(* IEC 61131-3 sources: volt/packages/volt-lsp-iec/test-corpus/awa-palletizer/Device/Plc Logic/Application/Library Manager/L_TW2P_TechModulesWindingTraversing, 72 files *)

(* ---- L_TW2P_ADAPTSPDCTRLGAINMODE.dut ---- *)
TYPE L_TW2P_ADAPTSPDCTRLGAINMODE :
(
	DIAMTOSQUARE := 0,
	DIAM := 1,
	INERTIA := 2
);
END_TYPE

(* ---- L_TW2P_DANCERCTRLSTOPMODE.dut ---- *)
TYPE L_TW2P_DANCERCTRLSTOPMODE :
(
	HALT := 0,
	MOVEABS := 1,
	MOVEREL := 2,
	MOVEABSSHORTESTWAY := 3,
	STOPVELOCITYMASTER := 4
);
END_TYPE

(* ---- L_TW2P_DANCERLIMITMODE.dut ---- *)
TYPE L_TW2P_DANCERLIMITMODE :
(
	AUTOMATIC := 0,
	SCPARDANCERLIMITS := 1,
	TEACHEDDANCERLIMITS := 2
);
END_TYPE

(* ---- L_TW2P_PERSISTENTVARWINDER.dut ---- *)
TYPE L_TW2P_PERSISTENTVARWINDER :
STRUCT
	LRDIAM : LREAL;
	LRMATERIALCOUNTER : LREAL;
	LIREVCOUNTER : LINT;
	LRREVCOUNTERRESIDUAL : LREAL;
	XUPPERPOSTEACHED : BOOL;
	XLOWERPOSTEACHED : BOOL;
	LRDANCERUPPERLIMIT : LREAL;
	LRDANCERLOWERLIMIT : LREAL;
END_STRUCT
END_TYPE

(* ---- L_TW2P_RESETICTRLMODE.dut ---- *)
TYPE L_TW2P_RESETICTRLMODE :
(
	INSTANT := 0,
	RAMP := 1
);
END_TYPE

(* ---- L_TW2P_SCAP_TM_WINDER.dut ---- *)
TYPE L_TW2P_SCAP_TM_WINDER :
STRUCT
	AP_XSETVELOFFSET : BOOL;
	AP_LRVELOFFSET : LREAL;
	AP_XSETTRQOFFSET : BOOL;
	AP_LRSETTRQOFFSET : LREAL;
	AP_XSETVELOFFSETDIAMCACL : BOOL;
	AP_LRVELOFFSETDIAMCACL : LREAL;
	AP_XSETSPEEDPOINTDIAMCALC : BOOL;
	AP_LRSETSPEEDPOINTDIAMCALC : LREAL;
	AP_XSETSPEEDPOINT : BOOL;
	AP_LRSETSPEEDPOINT : LREAL;
	AP_XVIRTUALRATEDSPEED : BOOL;
	AP_LRVIRTUALRATEDSPEED : LREAL := 4000;
	AP_XVIRTUALRATEDTORQUE : BOOL;
	AP_LRVIRTUALRATEDTORQUE : LREAL := 100;
END_STRUCT
END_TYPE

(* ---- L_TW2P_SCAP_TM_WINDERDANCERCTRLBASE.dut ---- *)
TYPE L_TW2P_SCAP_TM_WINDERDANCERCTRLBASE :
STRUCT
	AP_XSETDANCERCTRLOUTGAIN : BOOL;
	AP_LRSETDANCERCTRLOUTGAIN : LREAL;
	AP_XSETDANCERCTRLOUTRESETTIME : BOOL;
	AP_LRSETDANCERCTRLOUTRESETTIME : LREAL;
	AP_XSETDANCERCTRLOUTRATETIME : BOOL;
	AP_LRSETDANCERCTRLOUTRATETIME : LREAL;
	AP_WPIDMODE : WORD;
END_STRUCT
END_TYPE

(* ---- L_TW2P_SCAP_TM_WINDERDANCERCTRLSTATE.dut ---- *)
TYPE L_TW2P_SCAP_TM_WINDERDANCERCTRLSTATE :
STRUCT
	AP_XSETTRQPOINT : BOOL;
	AP_LRSETTRQPOINT : LREAL;
END_STRUCT
END_TYPE

(* ---- L_TW2P_SCAP_TM_WINDERTENSIONCTRLBASE.dut ---- *)
TYPE L_TW2P_SCAP_TM_WINDERTENSIONCTRLBASE :
STRUCT
	AP_XSETACCCOMPTRQ : BOOL;
	AP_LRACCCOMPTRQ : LREAL;
	AP_XSETTRQPOINT : BOOL;
	AP_LRSETTRQPOINT : LREAL;
	AP_XSETUPPERSPEEDLIMIT : BOOL;
	AP_LRSETUPPERSPEEDLIMIT : LREAL;
	AP_XSETLOWERSPEEDLIMIT : BOOL;
	AP_LRSETLOWERSPEEDLIMIT : LREAL;
END_STRUCT
END_TYPE

(* ---- L_TW2P_SCAP_TM_WINDERTENSIONCTRLSTATE.dut ---- *)
TYPE L_TW2P_SCAP_TM_WINDERTENSIONCTRLSTATE :
STRUCT
	AP_XSETTENSIONCTRLOUTGAIN : BOOL;
	AP_LRSETTENSIONCTRLOUTGAIN : LREAL;
	AP_XSETTENSIONCTRLOUTRESETTIME : BOOL;
	AP_LRSETTENSIONCTRLOUTRESETTIME : LREAL;
	AP_XSETTENSIONCTRLOUTRATETIME : BOOL;
	AP_LRSETTENSIONCTRLOUTRATETIME : LREAL;
	AP_XSETFRICCOMPREELSPEED : BOOL;
	AP_LRSETFRICCOMPREELSPEED : LREAL;
	AP_WPIDMODE : WORD;
END_STRUCT
END_TYPE

(* ---- L_TW2P_SCAP_WINDERDANCERCTRLBASE.dut ---- *)
TYPE L_TW2P_SCAP_WINDERDANCERCTRLBASE :
STRUCT
END_STRUCT
END_TYPE

(* ---- L_TW2P_SCAP_WINDERDANCERCTRLSTATE.dut ---- *)
TYPE L_TW2P_SCAP_WINDERDANCERCTRLSTATE :
STRUCT
END_STRUCT
END_TYPE

(* ---- L_TW2P_SCAP_WINDERTENSIONCTRLBASE.dut ---- *)
TYPE L_TW2P_SCAP_WINDERTENSIONCTRLBASE :
STRUCT
END_STRUCT
END_TYPE

(* ---- L_TW2P_SCAP_WINDERTENSIONCTRLSTATE.dut ---- *)
TYPE L_TW2P_SCAP_WINDERTENSIONCTRLSTATE :
STRUCT
END_STRUCT
END_TYPE

(* ---- L_TW2P_SCPAR_TM_WINDER.dut ---- *)
TYPE L_TW2P_SCPAR_TM_WINDER :
STRUCT
	LRLINEJERK : LREAL := 10000;
	LRJOGLINEACC : LREAL := 100;
	LRJOGLINEDEC : LREAL := 100;
	LRJOGLINEVEL : LREAL := 10;
	LRSYNCLINEACC : LREAL := 100;
	LRSYNCLINEDEC : LREAL := 100;
	LRWEBBREAKWINDOW : LREAL := 0.1;
	LRMAXDIAM : LREAL := 180;
	LRMINDIAM : LREAL := 50;
	RFILTTIMEDIAM : REAL := 0.05;
	LRDIAMCALCREGULARDIST : LREAL := 1;
	LRDIAMCALCREDUCEDDIST : LREAL := 0.1;
	ALRADAPTDIAMX : ARRAY [1..9] OF LREAL := [0, 100, 200, 300, 400, 500, 600, 700, 800];
	ALRADAPTDIAMY : ARRAY [1..9] OF LREAL := [0, 100, 200, 300, 400, 500, 600, 700, 800];
	LRTENSCURVECTRLSCALED : LREAL := 0;
	LRTENSCURVESTARTDIAMSCALED : LREAL := 0;
	LRLINEVELREF : LREAL := 1000;
	LRMINLINEVEL : LREAL := 1;
	RFILTTIMEMATERIALCOUNTER : REAL := 0.0;
	LRSETMATERIALPOS : LREAL;
	LRMAXWNDSPD : LREAL := 100;
	LRHYSTLINESTANDSTILL : LREAL;
	EDIAMCALCVALUESOURCE : MC_SOURCE;
	XLINEVELDIAMCALC : BOOL;
	LRTARGETMATERIALCOUNTER : LREAL;
	LRDIAMCHANGERAMP : LREAL := 0.0;
	LRDIAMCHANGELIMIT : LREAL := 0.0;
END_STRUCT
END_TYPE

(* ---- L_TW2P_SCPAR_TM_WINDERDANCERCTRLBASE.dut ---- *)
TYPE L_TW2P_SCPAR_TM_WINDERDANCERCTRLBASE :
STRUCT
	LRDANCERPOSRAMP : LREAL := 1;
	LRDANCERPOSCTRLGAIN : LREAL := 1;
	LRDANCERPOSCTRLRESETTIME : LREAL := 0;
	ERESETICTRLMODE : L_TW2P_ResetICtrlMode;
	LRDANCERPOSCTRLLIMITPOS : LREAL := 1;
	LRDANCERPOSCTRLLIMITNEG : LREAL := -1;
	LRDANCERMAXPOSSCALED : LREAL := 0.95;
	LRDANCERMINPOSSCALED : LREAL := -0.95;
	XTEACHDANCERLIMITS : BOOL := FALSE;
	LRDANCERUPPERLIMIT : LREAL := 10000000;
	LRDANCERLOWERLIMIT : LREAL := 0;
	LRDANCERMATERIALLENGTH : LREAL := 0;
	LRDANCERINPOSWINDOWSCALED : LREAL := 0.2;
	RFILTTIMEACTDANCERPOSIN : REAL := 0.005;
	RFILTTIMEACTDANCERVELCOMP : REAL := 0;
	WWEBBREAKMODE : WORD := 1;
END_STRUCT
END_TYPE

(* ---- L_TW2P_SCPAR_TM_WINDERDANCERCTRLSTATE.dut ---- *)
TYPE L_TW2P_SCPAR_TM_WINDERDANCERCTRLSTATE :
STRUCT
	DWSELECTTENSCURVE : DWORD := 0;
	ALRTENSCURVE : ARRAY [1..65] OF LREAL;
	RFILTTIMEACCSPD : REAL := 0.005;
	LRACCCMPSDEADBANDTRQSCALED : LREAL := 0.1;
	LRACCCMPSGAINACC : LREAL := 1.05;
	LRACCCMPSGAINDEC : LREAL := 0.95;
	LRCONSTMINERTIA : LREAL := 1;
	LRMAXMINERTIA : LREAL := 10;
	RFILTTIMEIDENTMINERTIASPD : REAL := 0.01;
	RFILTTIMEIDENTMINERTIATRQ : REAL := 0.005;
	LRIDENTMINERTIAMAXSPDSCALED : LREAL := 0.2;
	LRIDENTMINERTIAMAXTRQSCALED : LREAL := 0.2;
	EADAPTSPDCTRLGAINMODE : L_TW2P_AdaptSpdCtrlGainMode := 2;
	LRADAPTSPDCTRLLOWLIMIT : LREAL := 0.2;
	ALRSPDCTRLGAINADAPTX : ARRAY [1..9] OF LREAL := [0, 0.2, 0.4, 0.6, 0.8, 1, 1.2, 1.4, 1.6];
	ALRSPDCTRLGAINADAPTY : ARRAY [1..9] OF LREAL := [0, 0.2, 0.4, 0.6, 0.8, 1, 1.2, 1.4, 1.6];
	LRREDUCEDGAINWINDOW : LREAL;
	LRREDUCEDGAIN : LREAL;
	EDANCERCTRLSTOPMODE : L_TW2P_DancerCtrlStopMode;
	EDANCERCTRLMODE : L_TW2P_WinderDancerControlMode := L_TW2P_WinderDancerControlMode.SpeedBased;
	LRIDENTDIAMVEL : LREAL := 10;
	LRIDENTDIAMACC : LREAL := 100;
	LRIDENTDIAMDEC : LREAL := 100;
	LRIDENTDIAMJERK : LREAL;
	WIDENTDIAMCALCCYCLES : WORD := 2;
	LRIDENTDIAMMAXDANCERPOS : LREAL := 0.5;
	LRIDENTDIAMSPDCTRLGAIN : LREAL := 0.5;
END_STRUCT
END_TYPE

(* ---- L_TW2P_SCPAR_TM_WINDERTENSIONCTRLBASE.dut ---- *)
TYPE L_TW2P_SCPAR_TM_WINDERTENSIONCTRLBASE :
STRUCT
	LRLINEVELOFFSETSCALED : LREAL := 0.1;
	LRTENSREF : LREAL := 50;
	LRTENSRAMP : LREAL := 50;
	RFILTTIMEWNDSPD : REAL := 0.01;
	RFILTTIMEACCSPD : REAL := 0.005;
	LRACCCMPSDEADBANDTRQSCALED : LREAL := 0.1;
	LRACCCMPSGAINACC : LREAL := 1.05;
	LRACCCMPSGAINDEC : LREAL := 0.95;
	LRCONSTMINERTIA : LREAL := 1;
	LRMAXMINERTIA : LREAL := 10;
	LRFRICCURVESTARTTRQ : LREAL := 0;
	LRFRICCURVEENDTRQ : LREAL := 0;
	RFILTTIMEFRICSETSPD : REAL := 0.01;
END_STRUCT
END_TYPE

(* ---- L_TW2P_SCPAR_TM_WINDERTENSIONCTRLSTATE.dut ---- *)
TYPE L_TW2P_SCPAR_TM_WINDERTENSIONCTRLSTATE :
STRUCT
	DWSELECTTENSCURVE : DWORD := 0;
	ALRTENSCURVE : ARRAY [1..65] OF LREAL;
	LRTENSCTRLGAIN : LREAL := 0;
	LRTENSCTRLRESETTIME : LREAL := 0;
	ERESETICTRLMODE : L_TW2P_ResetICtrlMode;
	LRTENSCTRLLIMITPOS : LREAL := L_UMTP_Math.gC_POSITIVE_LIMIT_32BIT;
	LRTENSCTRLLIMITNEG : LREAL := L_UMTP_Math.gC_NEGATIVE_LIMIT_32BIT;
	LRIDENTFRICMAXSPDSCALED : LREAL := 0.9;
	LRIDENTFRICACCDEC : LREAL := 1;
	RFILTTIMEIDENTFRICSPD : REAL := 0.0;
	RFILTTIMEIDENTFRICTRQ : REAL := 0.05;
	DWSELECTFRICCURVE : DWORD := 1;
	RFILTTIMEACTTENSIN : REAL := 0.005;
	LRACTTENSINGAIN : LREAL := 1;
	LRACTTENSINOFFSET : LREAL := 0;
	RFILTTIMEIDENTMINERTIASPD : REAL := 0.01;
	RFILTTIMEIDENTMINERTIATRQ : REAL := 0.005;
	LRIDENTMINERTIAMAXSPDSCALED : LREAL := 0.2;
	LRIDENTMINERTIAMAXTRQSCALED : LREAL := 0.2;
	EADAPTSPDCTRLGAINMODE : L_TW2P_AdaptSpdCtrlGainMode := 2;
	LRADAPTSPDCTRLLOWLIMIT : LREAL := 0.2;
	ALRSPDCTRLGAINADAPTX : ARRAY [1..9] OF LREAL := [0, 0.2, 0.4, 0.6, 0.8, 1, 1.2, 1.4, 1.6];
	ALRSPDCTRLGAINADAPTY : ARRAY [1..9] OF LREAL := [0, 0.2, 0.4, 0.6, 0.8, 1, 1.2, 1.4, 1.6];
	LRREDUCEDGAINWINDOW : LREAL;
	LRREDUCEDGAIN : LREAL;
	ETENSCTRLSTOPMODE : L_TW2P_TensionCtrlStopMode;
	ETENSCTRLMODE : L_TW2P_WinderTensionControlMode := L_TW2P_WinderTensionControlMode.TorqueBased;
	LRTENSINWINDOWSCALED : LREAL := 0.2;
END_STRUCT
END_TYPE

(* ---- L_TW2P_SCPAR_WINDERDANCERCTRLBASE.dut ---- *)
TYPE L_TW2P_SCPAR_WINDERDANCERCTRLBASE :
STRUCT
END_STRUCT
END_TYPE

(* ---- L_TW2P_SCPAR_WINDERDANCERCTRLSTATE.dut ---- *)
TYPE L_TW2P_SCPAR_WINDERDANCERCTRLSTATE :
STRUCT
END_STRUCT
END_TYPE

(* ---- L_TW2P_SCPAR_WINDERTENSIONCTRLBASE.dut ---- *)
TYPE L_TW2P_SCPAR_WINDERTENSIONCTRLBASE :
STRUCT
END_STRUCT
END_TYPE

(* ---- L_TW2P_SCPAR_WINDERTENSIONCTRLSTATE.dut ---- *)
TYPE L_TW2P_SCPAR_WINDERTENSIONCTRLSTATE :
STRUCT
END_STRUCT
END_TYPE

(* ---- L_TW2P_SCSF_TM_WINDER.dut ---- *)
TYPE L_TW2P_SCSF_TM_WINDER :
STRUCT
	MP_LRWNDVELREF : LREAL;
	MP_LRWNDSPEEDREF : LREAL;
	MP_LIREVCOUNTER : LINT;
	MP_LRREVCOUNTERRESIDUAL : LREAL;
	MP_LRAXISSPEED : LREAL;
	MP_XDIAMCALCULATED : BOOL;
	MP_LRSETDIAMUNFILTERED : LREAL;
	MP_LRSETDIAMADAPTED : LREAL;
	MP_LRSETDIAMSCALEDOUT : LREAL;
	MP_LRSETLINEVELSCALEDOUT : LREAL;
	MP_LRACTTOTALTRQSCALED : LREAL;
	MP_XLINESTANDSTILL : BOOL;
	MP_LRSETSPEEDPOINT : LREAL;
	MP_LRWNDSPEEDINTEGRATED : LREAL;
	MP_LRLINEVELINTEGRATED : LREAL;
	MP_LRDISTTOLINESTOP : LREAL;
	MP_LRTARGETMATERIALCOUNTERSTOPLINE : LREAL;
END_STRUCT
END_TYPE

(* ---- L_TW2P_SCSF_TM_WINDERDANCERCTRLBASE.dut ---- *)
TYPE L_TW2P_SCSF_TM_WINDERDANCERCTRLBASE :
STRUCT
	MP_LRDANCERPOSSCALED0TO1 : LREAL;
	MP_LRDANCERCOMPVELOUT : LREAL;
	MP_LRFILTDANCERCOMPVELOUT : LREAL;
	MP_LRFILTACTDANCERPOSSCALED : LREAL;
	MP_LRSETRAMPDANCERPOS : LREAL;
	MP_LRDANCERCTRLPOSOUT : LREAL;
	MP_LRPDANCERCTRLOUT : LREAL;
	MP_LRIDANCERCTRLOUT : LREAL;
	MP_LRDDANCERCTRLOUT : LREAL;
	MP_LRDANCERCTRLLINEVELOUT : LREAL;
	MP_LRDANCERCTRLOUTGAIN : LREAL;
	MP_LRDANCERCTRLOUTRESETTIME : LREAL;
	MP_LRDANCERCTRLOUTRATETIME : LREAL;
	MP_LRDANCERCTRLSCALEDOUT : LREAL;
END_STRUCT
END_TYPE

(* ---- L_TW2P_SCSF_TM_WINDERDANCERCTRLSTATE.dut ---- *)
TYPE L_TW2P_SCSF_TM_WINDERDANCERCTRLSTATE :
STRUCT
	MP_LRAXISTORQUE : LREAL;
	MP_LRSETTRQPOINT : LREAL;
	MP_LRACCCOMPTRQ : LREAL;
	MP_LRACCTRQSCALEDOUT : LREAL;
END_STRUCT
END_TYPE

(* ---- L_TW2P_SCSF_TM_WINDERTENSIONCTRLBASE.dut ---- *)
TYPE L_TW2P_SCSF_TM_WINDERTENSIONCTRLBASE :
STRUCT
	MP_LRTENSCURVEOUT : LREAL;
	MP_LRSETTENSPOINT : LREAL;
	MP_LRSETTENSTRQ : LREAL;
	MP_LRACCCOMPTRQ : LREAL;
	MP_LRSETFRICCOMPTRQ : LREAL;
	MP_LRSETTRQPOINT : LREAL;
	MP_LRSETUPPERSPEEDLIMIT : LREAL;
	MP_LRSETLOWERSPEEDLIMIT : LREAL;
	MP_LRAXISUPPERSPEEDLIMIT : LREAL;
	MP_LRAXISLOWERSPEEDLIMIT : LREAL;
	MP_LRAXISVEL : LREAL;
	MP_LRAXISTORQUE : LREAL;
	MP_LRSETTENSSCALEDOUT : LREAL;
	MP_LRSETTENSTRQSCALEDOUT : LREAL;
	MP_LRSETFRICTRQSCALEDOUT : LREAL;
	MP_LRACCTRQSCALEDOUT : LREAL;
END_STRUCT
END_TYPE

(* ---- L_TW2P_SCSF_TM_WINDERTENSIONCTRLSTATE.dut ---- *)
TYPE L_TW2P_SCSF_TM_WINDERTENSIONCTRLSTATE :
STRUCT
	MP_LRFILTACTTENSIN : LREAL;
	MP_LRTENSCTRLOUT : LREAL;
	MP_LRPTENSCTRLOUT : LREAL;
	MP_LRITENSCTRLOUT : LREAL;
	MP_LRDTENSCTRLOUT : LREAL;
	MP_LRTENSCTRLOUTGAIN : LREAL;
	MP_LRTENSCTRLOUTRESETTIME : LREAL;
	MP_LRTENSCTRLOUTRATETIME : LREAL;
	MP_LRTENSCTRLOUTSCALED : LREAL;
	MP_LRSETTENSCTRLVALUE : LREAL;
	MP_LRACTTENSCTRLVALUE : LREAL;
	MP_LRACTTENSSCALED : LREAL := 0;
	MP_XSETTENSINTARGET : BOOL;
	MP_XACTTENSINTARGET : BOOL;
END_STRUCT
END_TYPE

(* ---- L_TW2P_SCSF_WINDERDANCERCTRLBASE.dut ---- *)
TYPE L_TW2P_SCSF_WINDERDANCERCTRLBASE :
STRUCT
END_STRUCT
END_TYPE

(* ---- L_TW2P_SCSF_WINDERDANCERCTRLSTATE.dut ---- *)
TYPE L_TW2P_SCSF_WINDERDANCERCTRLSTATE :
STRUCT
END_STRUCT
END_TYPE

(* ---- L_TW2P_SCSF_WINDERTENSIONCTRLBASE.dut ---- *)
TYPE L_TW2P_SCSF_WINDERTENSIONCTRLBASE :
STRUCT
END_STRUCT
END_TYPE

(* ---- L_TW2P_SCSF_WINDERTENSIONCTRLSTATE.dut ---- *)
TYPE L_TW2P_SCSF_WINDERTENSIONCTRLSTATE :
STRUCT
END_STRUCT
END_TYPE

(* ---- L_TW2P_TENSIONCTRLSTOPMODE.dut ---- *)
TYPE L_TW2P_TENSIONCTRLSTOPMODE :
(
	HALT := 0,
	MOVEABS := 1,
	MOVEREL := 2,
	MOVEABSSHORTESTWAY := 3,
	STOPVELOCITYMASTER := 4
);
END_TYPE

(* ---- L_TW2P_WINDERDANCERCONTROLMODE.dut ---- *)
TYPE L_TW2P_WINDERDANCERCONTROLMODE :
(
	SPEEDBASED := 1,
	VELOCITYMASTER := 2
);
END_TYPE

(* ---- L_TW2P_WINDERDANCERCTRLSTATEIN.dut ---- *)
TYPE L_TW2P_WINDERDANCERCTRLSTATEIN :
STRUCT
	XTEACHUPPERPOS : BOOL;
	XTEACHLOWERPOS : BOOL;
	XDANCERCTRL : BOOL;
	XRESETICTRL : BOOL;
	LRACTDANCERPOSIN : LREAL;
	LRSETDANCERPOSSCALED : LREAL;
	LRCTRLINFLUENCESCALED : LREAL;
	XACCCMPS : BOOL;
	LRMINERTIAADAPT : LREAL;
	XEXECUTEIDENTMINERTIA : BOOL;
	XEXECUTEIDENTDIAM : BOOL;
	XADAPTSPDCTRLGAIN : BOOL;
	LRADAPTSPDCTRLGAINFACTOR : LREAL;
END_STRUCT
END_TYPE

(* ---- L_TW2P_WINDERDANCERCTRLSTATEOUT.dut ---- *)
TYPE L_TW2P_WINDERDANCERCTRLSTATEOUT :
STRUCT
	XDANCERREACHEDSETPOS : BOOL;
	XDANCERMAXPOS : BOOL;
	XDANCERMINPOS : BOOL;
	LRACTDANCERPOSSCALED : LREAL;
	LRSETTENSCURVEOUT : LREAL;
	LRSETMINERTIAOUT : LREAL;
	LRIDENTMINERTIA : LREAL;
	LRSETSPDCTRLGAINADAPTOUT : LREAL;
END_STRUCT
END_TYPE

(* ---- L_TW2P_WINDERIN.dut ---- *)
TYPE L_TW2P_WINDERIN :
STRUCT
	MATERIALCOUNTERVALUES : L_MC1P_IAXIS_REF_MASTERVALUES;
	PERSISTENTVAR : L_TW2P_PersistentVarWinder;
	XMATERIALFEEDING : BOOL;
	XWINDINGDIRECTION : BOOL;
	XSETMATERIALCOUNTER : BOOL;
	XLOADDIAM : BOOL;
	LRLOADDIAM : LREAL;
	XHOLDDIAM : BOOL;
	XDIAMCALCREDUCED : BOOL;
	XWEBBREAKMONIT : BOOL;
	XJOGLINEPOS : BOOL;
	XJOGLINENEG : BOOL;
	XSYNCIN : BOOL;
	XTENSCURVE : BOOL;
	LRSETTENS : LREAL;
	LRSETLINEVEL : LREAL;
	LRSETLINEVELDIAMCALC : LREAL;
END_STRUCT
END_TYPE

(* ---- L_TW2P_WINDEROUT.dut ---- *)
TYPE L_TW2P_WINDEROUT :
STRUCT
	XWINDINGBUSY : BOOL;
	XSYNCHRONISED : BOOL;
	XACCDECSYNC : BOOL;
	XIDENTBUSY : BOOL;
	XIDENTDONE : BOOL;
	XUNWIND : BOOL;
	XWEBBREAK : BOOL;
	XHOLDDIAMACTIVE : BOOL;
	XDIAMMAX : BOOL;
	XDIAMMIN : BOOL;
	LRSETDIAMOUT : LREAL;
	LRMATERIALCOUNTER : LREAL;
	LRLIMITLINEVEL : LREAL;
	XVELOCITYMASTERBUSY : BOOL;
	LRSETLINEVELOUT : LREAL;
	XLINESTOP : BOOL;
	XMATERIALCOUNTERAXISVALID : BOOL;
END_STRUCT
END_TYPE

(* ---- L_TW2P_WINDERTENSIONCONTROLMODE.dut ---- *)
TYPE L_TW2P_WINDERTENSIONCONTROLMODE :
(
	TORQUEBASED := 0,
	SPEEDBASED := 1,
	VELOCITYMASTER := 2
);
END_TYPE

(* ---- L_TW2P_WINDERTENSIONCTRLSTATEIN.dut ---- *)
TYPE L_TW2P_WINDERTENSIONCTRLSTATEIN :
STRUCT
	XWINDINGDIRECTIONSTANDSTILL : BOOL;
	XTENSCTRL : BOOL;
	XFRICCMPS : BOOL;
	XACCCMPS : BOOL;
	LRMINERTIAADAPT : LREAL;
	XRESETPICTRL : BOOL;
	XRESETICTRL : BOOL;
	LRACTTENSIN : LREAL := 0;
	LRSETFRICADAPT : LREAL;
	LRCTRLINFLUENCESCALED : LREAL := 0;
	XEXECUTEIDENTFRIC : BOOL;
	XEXECUTEIDENTMINERTIA : BOOL;
	XADAPTSPDCTRLGAIN : BOOL;
	LRADAPTSPDCTRLGAINFACTOR : LREAL;
	LRMAXMINERTIA : LREAL;
END_STRUCT
END_TYPE

(* ---- L_TW2P_WINDERTENSIONCTRLSTATEOUT.dut ---- *)
TYPE L_TW2P_WINDERTENSIONCTRLSTATEOUT :
STRUCT
	XCONSTANTTENSION : BOOL;
	XWNDSPDLIMIT : BOOL;
	LRSETMINERTIAOUT : LREAL;
	XTENSINTARGET : BOOL;
	LRIDENTMINERTIA : LREAL;
	LRSETSPDCTRLGAINADAPTOUT : LREAL;
END_STRUCT
END_TYPE

(* ---- GETBOOLEANPROPERTY.pou ---- *)
FUNCTION GETBOOLEANPROPERTY : BOOL
VAR_INPUT
	STKEY : WSTRING;
END_VAR
END_FUNCTION

(* ---- GETCOMPANY.pou ---- *)
FUNCTION GETCOMPANY : WSTRING
END_FUNCTION

(* ---- GETNUMBERPROPERTY.pou ---- *)
FUNCTION GETNUMBERPROPERTY : DINT
VAR_INPUT
	STKEY : WSTRING;
END_VAR
END_FUNCTION

(* ---- GETTEXTPROPERTY.pou ---- *)
FUNCTION GETTEXTPROPERTY : WSTRING
VAR_INPUT
	STKEY : WSTRING;
END_VAR
END_FUNCTION

(* ---- GETTEXTPROPERTY2.pou ---- *)
FUNCTION GETTEXTPROPERTY2 : POINTER TO WSTRING
VAR_INPUT
	STKEY : WSTRING;
END_VAR
END_FUNCTION

(* ---- GETTITLE.pou ---- *)
FUNCTION GETTITLE : WSTRING
END_FUNCTION

(* ---- GETVERSION.pou ---- *)
FUNCTION GETVERSION : VERSION
END_FUNCTION

(* ---- GETVERSIONPROPERTY.pou ---- *)
FUNCTION GETVERSIONPROPERTY : VERSION
VAR_INPUT
	STKEY : WSTRING;
END_VAR
END_FUNCTION

(* ---- L_TW2P_CALCIDENDIAMETERBASE.pou ---- *)
FUNCTION L_TW2P_CALCIDENDIAMETERBASE : LREAL
VAR_IN_OUT
	LRLINEDIST : LREAL;
	LRDIAMCALCDIST : LREAL;
END_VAR
END_FUNCTION

(* ---- L_TW2P_CALCIDENDIAMETERSTATE.pou ---- *)
FUNCTION L_TW2P_CALCIDENDIAMETERSTATE : LREAL
VAR_IN_OUT
	LRDANCERPOSSTART : LREAL;
	LRDANCERPOSEND : LREAL;
	LRDIAMCALCDIST : LREAL;
	LRDANCERMATERIALLENGTH : LREAL;
END_VAR
END_FUNCTION

(* ---- L_TW2P_CONVERTPOSTOMODULOPOS.pou ---- *)
FUNCTION L_TW2P_CONVERTPOSTOMODULOPOS : LREAL
VAR_INPUT
	LRPOS : LREAL;
	LRPERIOD : LREAL;
END_VAR
VAR_OUTPUT
	DIREVCOUNTER : DINT;
END_VAR
END_FUNCTION

(* ---- L_TW2P_CONVERTPOSTOMODULOPOSEXTENDED.pou ---- *)
FUNCTION L_TW2P_CONVERTPOSTOMODULOPOSEXTENDED : LREAL
VAR_INPUT
	LRPOS : LREAL;
	LRPERIOD : LREAL;
END_VAR
VAR_OUTPUT
	DIREVCOUNTER : DINT;
END_VAR
END_FUNCTION

(* ---- L_TW2P_GETTASKCYCLE.pou ---- *)
FUNCTION L_TW2P_GETTASKCYCLE : LREAL
END_FUNCTION

(* ---- L_TW2P_HLPDELTAVELTIMEEXTENDED.pou ---- *)
FUNCTION L_TW2P_HLPDELTAVELTIMEEXTENDED : BOOL
VAR_INPUT
	LRVELSTART : LREAL;
	LRACCSTART : LREAL;
	LRMAXACC : LREAL;
	LRMAXJERK : LREAL;
END_VAR
VAR_OUTPUT
	LRTIME : LREAL;
	LRDIST : LREAL;
END_VAR
END_FUNCTION

(* ---- GLOBALTEXTLIST.pou ---- *)
FUNCTION_BLOCK GLOBALTEXTLIST
VAR
	M_TEXTLISTFILE : STRING(255);
	_STNAMESPACE : STRING;
END_VAR
END_FUNCTION_BLOCK

(* ---- L_TW2P_DANCERSIMULATOR.pou ---- *)
FUNCTION_BLOCK L_TW2P_DANCERSIMULATOR
VAR_INPUT
	XENABLE : BOOL;
	XINVERT : BOOL;
	LRSETSPEED : LREAL;
	LRSETLINEVEL : LREAL;
	LRSETDIAM : LREAL := 120;
	LRMINDIAM : LREAL := 100;
	LRMATERIALDANCELENGHT : LREAL := 200;
	LRDANCERUPPERLIMIT : LREAL := 1;
	LRDANCERLOWERLIMIT : LREAL := -1;
	LRTASKCYCLE : LREAL := 0.001;
END_VAR
VAR_OUTPUT
	XBUSY : BOOL;
	LRSETDANCERPOSOUT : LREAL;
END_VAR
VAR
	_XENABLEOLD : BOOL;
	_LRDIAM : LREAL := 120;
	_LRMATERIALDANCELENGHT : LREAL := 200;
	_LRDANCERUPPERLIMIT : LREAL := 1;
	_LRDANCERLOWERLIMIT : LREAL := -1;
	_LRCALCCIRCUMFERENCEVEL : LREAL;
	_LRDELTALINEVEL : LREAL;
	_LRCALCMATIALDANCERLENGT : LREAL;
	_LRDANCERPOSSCALED : LREAL;
	_LRDANCERPOSSCALED2 : LREAL;
	_LRTASKCYCLE : LREAL := 0.001;
END_VAR
END_FUNCTION_BLOCK

(* ---- L_TW2P_MATERIALLENGTHCOUNTERFROMPOS.pou ---- *)
FUNCTION_BLOCK L_TW2P_MATERIALLENGTHCOUNTERFROMPOS
VAR_INPUT
	XENABLE : BOOL;
	LRACTPOSIN : LREAL;
	WFILTERDEPTH : WORD := 0;
	LRCYCLELENGTH : LREAL := 360;
	LRSETFEEDCONSTANT : LREAL := 360;
	XSETMATERIALCOUNTER : BOOL;
	LRSETMATERIALPOS : LREAL;
END_VAR
VAR_OUTPUT
	XBUSY : BOOL;
	XERROR : BOOL;
	EERRORID : L_IE1P_Error;
	LRMATERIALCOUNTER : LREAL;
	LRREVCOUNTER : LREAL;
	LIREVCOUNTER : LINT;
	LIREVCOUNTERMID : LINT;
	LRREVCOUNTERRESIDUAL : LREAL;
END_VAR
VAR_IN_OUT
	LIREVCOUNTERRETAIN : LINT;
	LRREVCOUNTERRESIDUALRETAIN : LREAL;
END_VAR
VAR
	WSTATE : WORD;
	XENABLE_OLD : BOOL;
	XSETMATERIALCOUNTER_OLD : BOOL;
	LRSTARTPOS_INT : LREAL;
	LRACTPOSIN_INT : LREAL;
	LIREVCOUNTER_OLD : LINT;
	LRREVCOUNTER_INT : LREAL;
	LIREVCOUNTERMID_OLD : LINT;
	LRREVCOUNTERMID_INT : LREAL;
	XERRORRECIVEDLIMIT : BOOL;
	LRREVCOUNTERRESIDUAL_OFFSET : LREAL;
	LRACTPOSIN_OLD : LREAL;
	C_LRLINTMAXVALUEPOS : LREAL := 2#111111111111111111111111111111111111111111111111111111111111111;
	C_LRLINTMAXVALUENEG : LREAL := -2#111111111111111111111111111111111111111111111111111111111111111;
END_VAR
END_FUNCTION_BLOCK

METHOD CALL_CALCMATERAILCOUNTER
END_METHOD

METHOD CALL_ERRORHANDLER
END_METHOD

METHOD CALL_OUTPUT
END_METHOD

METHOD CALL_RESETCOMMANDS
END_METHOD

METHOD CALL_RESETOUTPUT
END_METHOD

(* ---- L_TW2P_MATERIALLENGTHCOUNTERFROMVEL.pou ---- *)
FUNCTION_BLOCK L_TW2P_MATERIALLENGTHCOUNTERFROMVEL
VAR_INPUT
	XENABLE : BOOL;
	LRACTVELIN : LREAL;
	RFILTERTIME : REAL := 0.0;
	XSETMATERIALCOUNTER : BOOL;
	LRSETMATERIALPOS : LREAL;
END_VAR
VAR_OUTPUT
	XBUSY : BOOL;
	XWARNING : BOOL;
	EERRORID : L_IE1P_Error;
	LRMATERIALCOUNTER : LREAL;
END_VAR
VAR_IN_OUT
	LRSETMATERIALPOSRETAIN : LREAL;
END_VAR
VAR
	WSTATE : WORD;
	XENABLE_OLD : BOOL;
	XSETMATERIALCOUNTER_OLD : BOOL;
	LRTASKCYCLE : LREAL;
	LIPOS_INT : LINT;
	LIDELTAPOS_INT : LINT;
	LIPOS_OLD : LINT;
	LIIDX : LINT;
	LRMATERIALCOUNTERCOUNTER_INT : LREAL;
	LRMATERIALOFFSET_INT : LREAL;
	FB_PT1FILTER : L_USPP_PT1Filter;
END_VAR
END_FUNCTION_BLOCK

METHOD CALL_CALCMATERAILCOUNTER
END_METHOD

METHOD CALL_ERRORHANDLER
END_METHOD

METHOD CALL_FBMETHODS
END_METHOD

METHOD CALL_FB_PT1FILTER
END_METHOD

METHOD CALL_OUTPUT
END_METHOD

METHOD CALL_RESETCOMMANDS
END_METHOD

METHOD CALL_RESETOUTPUT
END_METHOD

METHOD CALL_STATEMACHINE
END_METHOD

(* ---- L_TW2P_RAMPDIAMETER.pou ---- *)
FUNCTION_BLOCK L_TW2P_RAMPDIAMETER
VAR_INPUT
	LRDIAMCHANGERAMP : LREAL;
	LRSETDIAM : LREAL;
	XLOADDIAM : BOOL;
END_VAR
VAR_OUTPUT
	XACTIVE : BOOL;
	LRSETDIAMOUT : LREAL;
END_VAR
VAR
	_XINITDONE : BOOL;
	_XLOADRAMPGENDONE : BOOL;
	FBRAMPGENERATOR : L_MC1P_RampGenerator;
END_VAR
END_FUNCTION_BLOCK

(* ---- L_TW2P_TM_WINDER.pou ---- *)
FUNCTION_BLOCK L_TW2P_TM_WINDER EXTENDS L_TB2P_TM_MotionControl
VAR_IN_OUT
	PERSISTENTVAR : L_TW2P_PersistentVarWinder;
END_VAR
VAR
	PINPUTWINDER : POINTER TO L_TW2P_WinderIn;
	POUTPUTWINDER : POINTER TO L_TW2P_WinderOut;
	XWINDINGBUSY : BOOL;
	XSYNCHRONISED : BOOL;
	XACCDECSYNC : BOOL;
	XIDENTBUSY : BOOL;
	XIDENTDONE : BOOL;
	XUNWIND : BOOL;
	XWEBBREAK : BOOL;
	XHOLDDIAMACTIVE : BOOL;
	XDIAMMAX : BOOL;
	XDIAMMIN : BOOL;
	LRSETDIAMOUT : LREAL;
	LRMATERIALCOUNTER : LREAL;
	LRLIMITLINEVEL : LREAL;
	XVELOCITYMASTERBUSY : BOOL;
	LRSETLINEVELOUT : LREAL;
	XLINESTOP : BOOL;
	LRTARGETMATERIALCOUNTERSTOPLINE_INT : LREAL;
	LRDISTTOLINESTOP_INT : LREAL;
	LRSETLINEVEL_INT : LREAL;
	LRSETLINEVELOUT_INT : LREAL;
	WWINDERSTOPMODE : WORD;
	XSELVELOCITYMASTERMODE_LOCK : BOOL;
	XVELOCITYMASTER_INT : BOOL;
	XUSEVIRTUALMODE_INT : BOOL;
	XWINDINGDIRECTIONSTANDSTILL_INT : BOOL := FALSE;
	XTRIMLINEPOS_INT : BOOL;
	XTRIMLINENEG_INT : BOOL;
	AP_XSETTRQOFFSET_INT : BOOL;
	AP_LRSETTRQOFFSET_INT : LREAL;
	AP_XSETVELOFFSET_INT : BOOL;
	AP_LRVELOFFSET_INT : LREAL;
	XLINEVELDIAMCALC_INT : BOOL;
	LRSETLINEVELDIAMCALC_INT : LREAL;
	XINVERTDIRECTION : BOOL;
	LRREELSPEEDINTEGRATE : LREAL;
	LRHALTDEC_INT : LREAL;
	LRHALTJERK_INT : LREAL;
	XLINESTANDSTILL_INT : BOOL;
	XFUNCTIONCANENABLE_INT : BOOL;
	XFUNCTIONHALTABORT_INT : BOOL;
	XUNWIND_OLD : BOOL;
	LRSETDIAMOUT_OLD : LREAL;
	XLOADDIAM_OLD : BOOL;
	XSYNCIN_OLD : BOOL;
	XERRORINVALIDINVERTER : BOOL;
	XWARNININVALIDINVERTER : BOOL;
	XWARNINGAXISNOTHOMED : BOOL;
	XWARNINGHOMINGBLOCKED : BOOL;
	XWARNINGDIRECTIONDISABLED_WINDING : BOOL;
	XWARNINGDIRECTIONDISABLED_SYNCLINEVEL : BOOL;
	XWARNINGDIRECTIONDISABLED_JOGLINEVEL : BOOL;
	XWARNINGDIRECTIONDISABLED_VELCITYMASTER : BOOL;
	DISETLOWERSPEEDLIMIT : DINT;
	DISETUPPERSPEEDLIMIT : DINT;
	DIOFFSETTORQUE : DINT;
	LRVIRTUALRATEDSPEED : LREAL;
	LRVIRTUALRATEDTORQUE : LREAL;
	LRVIRTUALRATEDTORQUEINV : LREAL;
	LRREFERENCEMOTORREELSPEED : LREAL := 0;
	LRREFERENCEREELSPEEDWINDER : LREAL := 0;
	LRREFERENCETORQUEWINDER : LREAL := 0;
	LRREFERENCETORQUEWINDERINV : LREAL;
	LRREFERENCEMOTORTORQUE : LREAL := 0;
	LRFEEDCONSTANT : LREAL;
	LRFEEDCONSTANT_ABS : LREAL;
	LRFEEDCONSTANTINV : LREAL;
	LRFEEDCONSTANTINV_ABS : LREAL;
	LRCYCLELENGTH_INV : LREAL;
	LRCYCLELENGTH : LREAL;
	LRGEARNUMERATOR : LREAL;
	LRGEARDENOMINATOR : LREAL;
	DWGEARDENOMINATOR_LOCK : DWORD;
	DWGEARNUMERATOR_LOCK : DWORD;
	XIDENTDIAMACTIVE : BOOL;
	LRREADAXISREELSPEED : LREAL;
	LRDIAMCALCREELSPEED : LREAL;
	LRCIRCUMFERENCE : LREAL;
	LRCIRCUMFERENCE_INV : LREAL;
	XSPEEDLIMITENABLED : BOOL;
	XDECOUPLINGLIMITREELSPEED : BOOL;
	XDCALCDISTANCEINIT : BOOL;
	WWINDERID : WORD;
	LRMINLINEVEL : LREAL;
	LRSETWNDSPEEDUPPERLIMIT : LREAL;
	LRSETWNDSPEEDLOWERLIMIT : LREAL;
	LRSETSPEEDCTRLGAINADAPT : LREAL := 1;
	LRSETSPEEDOFFSET : LREAL := 0;
	XTRIGGERCALCDIAM : BOOL;
	XTRIGGERCALCDIAM_OLD : BOOL;
	WNUMOFAXIS : WORD;
	XMATERIALCOUNTERAXISVALID : BOOL := FALSE;
	ETMSTATE_EXITSELECTMODE : L_TB2P_States := 2;
	ECONTROLMODECAMEFROM : L_MC1P_ControlMode;
	XWAITNEXTCYCLEFORSETCONTROLERMODE : BOOL;
	XSELECTCSVACTIVE_INT : BOOL;
	XSELECTCSPACTIVE_INT : BOOL;
	XSELECTCSTACTIVE_INT : BOOL;
	AP_XSETCONTROLLERMODE : BOOL;
	XSTOPMODEVIAHALT_INT : BOOL;
	PPARWINDER : POINTER TO L_TW2P_scPar_TM_Winder;
	XNEWREQUESTRESTARTFROMEXTERNAL : BOOL;
	XWEBBREAKEXT : BOOL := FALSE;
	LRPICTRLINTVALUE : LREAL := 0;
	XPICTRLLOADINTVALUE : BOOL := FALSE;
	XENABLETRQOFFSET : BOOL;
	LRACTTOTALTORQUE : LREAL;
	LRSETTORQUEOFFSET : LREAL := 0;
	LRSETTOTALTORQUE : LREAL;
	LRSETMOTORTORQUE : LREAL;
	LRACTMOTORTORQUE : LREAL;
	LRSETTOTALVELOCITY : LREAL;
	LRSETSPEEDTOTAL : LREAL;
	XDANCERMATERIALLENGTH : BOOL;
	LRACTDANCERLINEVELCOMP : LREAL := 0;
	LRVARMINERTIASCALED : LREAL;
	LRWNDVELREF : LREAL;
	LRSETPOSITION_OLD : LREAL;
	XDIAMCALCULATED_INT : BOOL;
	LRDIAMETERUNFILTERED_INT : LREAL;
	XTMHALT_INT : BOOL;
	XTMHALT_OLD : BOOL;
	LRMASTERVELFORTRANSITION : LREAL;
	LRMASTERVELFORTRANSITIONLINEJOGGING : LREAL;
	IACTMASTERDIRECTIONTMP : INT;
	IACTMASTERDIRECTIONLINEJOGGING : INT;
	FB_READPARAMETER : MC_ReadParameter;
	FB_READHALTDEC : MC_ReadParameter := STRUCT(ParameterNumber := 186);
	FB_READHALTJERK : MC_ReadParameter := STRUCT(ParameterNumber := 187);
	FB_READMACHINEDATA : L_MC1P_ReadmachineData;
	FB_FOLLOWVELOCITY : L_MC1P_ControlSetValues;
	FB_TORQUEOFFSET : L_MC1P_SetTorqueOffset;
	FB_HYSTERISIS : L_UMTP_Hysteresis;
	FB_SETCONTROLLERMODE : L_MC1P_SetControlMode;
	FB_TORQUECONTROL : L_MC1P_TorqueControl;
	L_MB1P_CURVESETDIAMETER : L_USPP_Curve;
	L_MB1P_CALCDIAMETER1 : L_TB1P_CalcDiameter;
	FB_RAMPDIAMETER : L_TW2P_RampDiameter;
	L_MB1P_TENSIONCURVE1 : L_TB1P_TensionCurve;
	FB_RAMPGENERATOR1 : L_MC1P_RampGenerator;
	FB_WINDERSYNCHRONISELINE1 : L_TW2P_WinderSynchroniseLine;
	FM_WINDERJOGGING1 : L_TW2P_WinderJogging;
	WMATERIALLENGTHCOUNTERMODE : WORD;
	FB_MATERIALLENGTHCOUNTER : L_TW2P_MaterialLengthCounterFromVel;
	FB_MATERIALLENGTHCOUNTERPOS : L_TW2P_MaterialLengthCounterFromPos;
	FB_VELOCITYMASTER : L_TW2P_WinderVelocityMaster;
	XINVALIDRETAIN : BOOL;
	LRSETDIAMOUTRETAIN : LREAL;
	XMOVEABSEXECUTEWINDER_INT : BOOL;
	XMOVERELEXECUTEWINDER_INT : BOOL;
	XMOVEVELEXECUTEWINDER_INT : BOOL;
	LRPOS_DISTWINDER_INT : LREAL;
	LRVELWINDER_INT : LREAL;
	LRACCWINDER_INT : LREAL;
	LRDECWINDER_INT : LREAL;
	LRJERKWINDER_INT : LREAL;
	EDIRECTIONWINDER_INT : MC_DIRECTION;
	XLINEJOGGINGBUSY_INT : BOOL;
END_VAR
END_FUNCTION_BLOCK

METHOD CALL_ALLOCPOINTADR
END_METHOD

METHOD CALL_CALCCIRCUMFERENCE
END_METHOD

METHOD CALL_CTRLREQACTIVE : BOOL
END_METHOD

METHOD CALL_ERRORHANDLER
END_METHOD

METHOD CALL_FBHYSTERISIS
END_METHOD

METHOD CALL_FBMETHODS
END_METHOD

METHOD CALL_FBMETHODS_WND
END_METHOD

METHOD CALL_FB_MATERIALLENGTHCOUNTER
END_METHOD

METHOD CALL_FB_MATERIALLENGTHCOUNTER_INPUT
END_METHOD

METHOD CALL_FB_RAMPGENERATOR
END_METHOD

METHOD CALL_FB_READHALTDEC
END_METHOD

METHOD CALL_FB_READHALTJERK
END_METHOD

METHOD CALL_FB_READPARAMETER
END_METHOD

METHOD CALL_FB_READMACHINEDATA
END_METHOD

METHOD CALL_FB_READMACHINEDATAMATCNTAXIS
END_METHOD

METHOD CALL_FB_SETCONTROLLERMODE
END_METHOD

METHOD CALL_FB_TORQUECONTROL
END_METHOD

METHOD CALL_FB_TORQUEOFFSET
END_METHOD

METHOD CALL_FB_VELOCITYMASTER
END_METHOD

METHOD CALL_FB_WINDERSYNCHRONISELINE
END_METHOD

METHOD CALL_FB_WNDCALCDIAMETER
END_METHOD

METHOD CALL_FB_WNDCALCDIAMETER_HOLDDIAMETER
END_METHOD

METHOD CALL_FB_WNDCALCDIAMETER_INPUT
END_METHOD

METHOD CALL_FB_WNDRAMPDIAMETER
END_METHOD

METHOD CALL_FM_WINDERJOGGING
END_METHOD

METHOD CALL_FIRSTCYCLE
END_METHOD

METHOD CALL_FOLLOWVELOCITY
END_METHOD

METHOD CALL_INITDONE
END_METHOD

METHOD CALL_INITROUTINE
END_METHOD

METHOD CALL_INTERNALCTRL
END_METHOD

METHOD CALL_LIMITLINEVEL
END_METHOD

METHOD CALL_LIMITEDINPUT
END_METHOD

METHOD CALL_OUTPUT
END_METHOD

METHOD CALL_READACTUALTORQUE
END_METHOD

METHOD CALL_READAXISREELSPEED
END_METHOD

METHOD CALL_REQUESTS_EXT
END_METHOD

METHOD CALL_RESETCOMMANDS
END_METHOD

METHOD CALL_RESETIDENTFBS
END_METHOD

METHOD CALL_RESETOUTPUT
END_METHOD

METHOD CALL_RESETPERSISTENTVARWINDER
END_METHOD

METHOD CALL_RESETWARNINGS
END_METHOD

METHOD CALL_SETPERSISTENTVARWINDER
END_METHOD

METHOD CALL_SETSPEEDPOINT
END_METHOD

METHOD CALL_SETTORQUE
END_METHOD

METHOD CALL_SETTORQUEOFFESET
END_METHOD

METHOD CALL_SETUNWINDSTATUS
END_METHOD

METHOD CALL_SETWINDERID
END_METHOD

METHOD CALL_STATEMACHINE
END_METHOD

METHOD CALL_TBCURVESETDIAMETER : LREAL
END_METHOD

METHOD CALL_WNDTENSIONCURVE
END_METHOD

METHOD CALL_WNDTENSIONCURVE_INPUT
END_METHOD

METHOD CALL_ABC_INPUT
END_METHOD

METHOD CALL_ABC_INPUT_PROFILEPARAMETER
END_METHOD

METHOD GET_ESTATE : L_TB2P_States
END_METHOD

METHOD GET_ETMSTATE : L_TB2P_States
END_METHOD

METHOD GET_LRACTMOTORTORQUE : LREAL
END_METHOD

METHOD GET_LRCALCDIAMDIST : LREAL
END_METHOD

METHOD GET_LRCALCDIAMLINESPEED : LREAL
END_METHOD

METHOD GET_LRCALCDIAMREELSPEED : LREAL
END_METHOD

METHOD GET_LRFEEDCONSTANT : LREAL
END_METHOD

METHOD GET_LRLOWERSPEEDLIMIT : LREAL
END_METHOD

METHOD GET_LRMOTORTORQUEREF : LREAL
END_METHOD

METHOD GET_LRREELSPEEDREF : LREAL
END_METHOD

METHOD GET_LRSETMOTORTORQUE : LREAL
END_METHOD

METHOD GET_LRSETSPEEDCTRLGAINADAPT : LREAL
END_METHOD

METHOD GET_LRSETTOTALTORQUE : LREAL
END_METHOD

METHOD GET_LRSETTOTALTRQ : LREAL
END_METHOD

METHOD GET_LRTASKCYCLE : LREAL
END_METHOD

METHOD GET_LRUPPERSPEEDLIMIT : LREAL
END_METHOD

METHOD GET_LRVARMINERTIASCALED : LREAL
END_METHOD

METHOD GET_LRWINDERTORQUEREF : LREAL
END_METHOD

METHOD GET_XCOMMUNICATION : BOOL
END_METHOD

METHOD GET_XDIAMWEBBREAKENABLE : BOOL
VAR_OUTPUT
	XUNIDIRECT : BOOL;
	XUNWINDACTIVE : BOOL;
END_VAR
END_METHOD

METHOD CALL_COUPLINGREELSPEEDLIMIT
END_METHOD

METHOD CALL_DECOUPLINGREELSPEEDLIMIT
END_METHOD

METHOD SET_ESTATE
VAR_INPUT
	IN : L_TB2P_States;
END_VAR
END_METHOD

METHOD SET_LRFEEDCONSTANT
VAR_INPUT
	LRIN : LREAL := 0;
END_VAR
END_METHOD

METHOD SET_LRPICTRLINTVALUE
VAR_INPUT
	LRIN : LREAL := 0;
END_VAR
END_METHOD

METHOD SET_LRREFERENCEMOTORTORQUE
VAR_INPUT
	LRIN : LREAL := 0;
END_VAR
END_METHOD

METHOD SET_LRREFERENCEREELSPEED
VAR_INPUT
	LRIN : LREAL := 0;
END_VAR
END_METHOD

METHOD SET_LRSPEEDOFFSET
VAR_INPUT
	LRIN : LREAL := 0;
END_VAR
END_METHOD

METHOD SET_LRTORQUEOFFSET
VAR_INPUT
	LRIN : LREAL := 0;
END_VAR
END_METHOD

METHOD SET_XPICTRLLOADINTVALUE
VAR_INPUT
	XIN : BOOL := FALSE;
END_VAR
END_METHOD

METHOD SET_XSPEEDLIMITENABLEDEXT
VAR_INPUT
	XIN : BOOL := TRUE;
END_VAR
END_METHOD

METHOD SET_XWEBBREAK
VAR_INPUT
	XIN : BOOL := FALSE;
END_VAR
END_METHOD

METHOD CALL_S000_CYCLIC
END_METHOD

METHOD CALL_S002_STANDBY
END_METHOD

METHOD CALL_S015_LINEJOGGING
END_METHOD

METHOD CALL_S020_SYNCLINEVEL
END_METHOD

METHOD CALL_S060_SELECTMODECSV
END_METHOD

METHOD CALL_S070_SELECTMODECST
END_METHOD

METHOD CALL_S071_VELOCITYMASTER
END_METHOD

METHOD CALL_S071_VELOCITYMASTER_STOP
END_METHOD

METHOD CALL_S123_SELECTMODECSP
END_METHOD

METHOD CALL_S996_STOP
END_METHOD

METHOD CALL_S999_ERROR
END_METHOD

METHOD CALL_T000_ALLSTATES
END_METHOD

METHOD CALL_T020_SYNCLINEVEL
END_METHOD

METHOD CALL_T071_VELOCITYMASTER
END_METHOD

METHOD CALL_S999_ERROR_OUT
END_METHOD

(* ---- L_TW2P_TM_WINDERDANCERCTRLBASE.pou ---- *)
FUNCTION_BLOCK L_TW2P_TM_WINDERDANCERCTRLBASE EXTENDS L_TW2P_TM_Winder
VAR_OUTPUT
	PPAR : POINTER TO L_TW2P_scPar_TM_WinderDancerCtrlState := ADR(scPar_int);
	PSF : POINTER TO L_TW2P_scSF_TM_WinderDancerCtrlState;
	PAP : POINTER TO L_TW2P_scAP_TM_WinderDancerCtrlState;
END_VAR
VAR
	PINPUTWINDERDANCER : POINTER TO L_TW2P_WinderDancerCtrlStateIn;
	POUTPUTWINDERDANCER : POINTER TO L_TW2P_WinderDancerCtrlStateOut;
	TM_WINDERDANCERCTRLBASECONFIG : L_TB2P_ModuleHandlerConfig;
	XDANCERREACHEDSETPOS : BOOL;
	XDANCERMAXPOS : BOOL;
	XDANCERMINPOS : BOOL;
	LRACTDANCERPOSSCALED : LREAL;
	LRSETTENSCURVEOUT : LREAL;
	XRESETTEACHDANCERPOS_INT : BOOL;
	XTEACHDANCERLIMITS_OLD : BOOL;
	XTEACHUPPERPOS_OLD : BOOL;
	XTEACHLOWERPOS_OLD : BOOL;
	XRESETICTRL_OLD : BOOL;
	LRDANCERPOSCTRLRESETTIME_STORE : LREAL;
	LRDEVIATION_STORE : LREAL;
	SCPAR_INT : L_TW2P_scPar_TM_WinderDancerCtrlState;
	XDANCERCONTROLACTIVE_INT : BOOL;
	LRSETREELSPEEDFRWCTRL : LREAL;
	LRSETREELSPEEDDEVIATION : LREAL;
	LRDANCERPOSCTRLOUTVEL : LREAL;
	LRDANCERPOSREF : LREAL;
	LRDANCERPOSSCALED0TO1 : LREAL;
	LRFILTACTDANCERPOS : LREAL;
	LRFILTACTDANCERPOSSCALED : LREAL;
	LRACTDANCERVEL : LREAL;
	XWARNING_DANCERLIMITSNOTTEACHED : BOOL;
	L_MB1P_RAMPGENERATORRESETICTRL : L_MC1P_RampGenerator;
	L_MB1P_DIFFERENTIATE1 : L_MC2P_Differentiate;
	L_MB1P_PROCESSCONTROLLER1 : L_CT1P_ProcessController;
	L_D94A_FILTERDANCERPOSIN : L_USPP_PT1Filter;
	L_D94A_FILTERLINEVELCOMP : L_USPP_PT1Filter;
	LRDANCERUPPERLIMIT_INT : LREAL;
	LRDANCERLOWERLIMIT_INT : LREAL;
	XUPPERPOSTEACHED : BOOL;
	XLOWERPOSTEACHED : BOOL;
	LRTEACHEDDANCERUPPERLIMIT_INT : LREAL;
	LRTEACHEDDANCERLOWERLIMIT_INT : LREAL;
END_VAR
END_FUNCTION_BLOCK

METHOD CALL_ALLOCPOINTADR
END_METHOD

METHOD CALL_CTRLREQACTIVE : BOOL
END_METHOD

METHOD CALL_ERRORHANDLER
END_METHOD

METHOD CALL_FBMETHODS
END_METHOD

METHOD CALL_FBMETHODS_WND
END_METHOD

METHOD CALL_FB_PROCESSCONTROLLER
END_METHOD

METHOD CALL_FB_RAMPGENERATOR
END_METHOD

METHOD CALL_FB_WNDCALCDIAMETER_INPUT
END_METHOD

METHOD CALL_FILTERDANCERPOSIN
END_METHOD

METHOD CALL_FILTERLINEVELCOMP
END_METHOD

METHOD CALL_FIRSTCYCLE
END_METHOD

METHOD CALL_INITROUTINE
END_METHOD

METHOD CALL_INTERNALCTRL
END_METHOD

METHOD CALL_OUTPUT
END_METHOD

METHOD CALL_OUTPUT_SF
END_METHOD

METHOD CALL_RAMPGENERATORRESETICTRL
END_METHOD

METHOD CALL_REQUESTS_EXT
END_METHOD

METHOD CALL_RESETCOMMANDS
END_METHOD

METHOD CALL_RESETOUTPUT
END_METHOD

METHOD CALL_RESETWARNINGS
END_METHOD

METHOD CALL_SDDIFFERENTIATE : BOOL
END_METHOD

METHOD CALL_SETSPEEDPOINT
END_METHOD

METHOD CALL_STATEMACHINE
END_METHOD

METHOD CALL_TEACHDANCER
END_METHOD

METHOD GET_LRACTDANCERCTRLOUT : LREAL
END_METHOD

METHOD GET_LRACTDANCERLINEVELCOMP : LREAL
END_METHOD

METHOD GET_LRACTDANCERVEL : LREAL
END_METHOD

METHOD GET_LRSPEEDFORWARDCTRL : LREAL
END_METHOD

METHOD GET_LRSPEEDSETPOINT : LREAL
END_METHOD

METHOD GET_LRVELSETPOINT : LREAL
END_METHOD

METHOD GET_XLOWERPOSTEACHED : BOOL
VAR_OUTPUT
	LRTEACHPOSLOWERLIMIT : LREAL;
END_VAR
END_METHOD

METHOD GET_XUPPERPOSTEACHED : BOOL
VAR_OUTPUT
	LRTEACHPOSUPPERLIMIT : LREAL;
END_VAR
END_METHOD

METHOD CALL_RESTDANCERTEACHPOS
END_METHOD

METHOD LOAD_LRDANCERLOWERLIMIT
VAR_INPUT
	LRIN : LREAL := 0;
END_VAR
END_METHOD

METHOD LOAD_LRDANCERUPPERLIMIT
VAR_INPUT
	LRIN : LREAL := 0;
END_VAR
END_METHOD

METHOD SET_ALRPROCESSCTRLXVALUES
VAR_INPUT
	ALRPROCESSCTRLXVALUES : ARRAY [1..5] OF LREAL;
END_VAR
END_METHOD

METHOD SET_ALRPROCESSCTRLYVALUES
VAR_INPUT
	ALRPROCESSCTRLYVALUES : ARRAY [1..5] OF LREAL;
END_VAR
END_METHOD

METHOD SET_LRPICTRLINTVALUE
VAR_INPUT
	LRIN : LREAL := 0;
END_VAR
END_METHOD

METHOD SET_LRPROCESSCTRLACC
VAR_INPUT
	LRPROCESSCTRLACC : LREAL := 0.0;
END_VAR
END_METHOD

METHOD SET_LRPROCESSCTRLDEC
VAR_INPUT
	LRPROCESSCTRLDEC : LREAL := 0.0;
END_VAR
END_METHOD

METHOD SET_LRPROCESSCTRLGAINADAPT
VAR_INPUT
	LRPROCESSCTRLGAINADAPT : LREAL := 1;
END_VAR
END_METHOD

METHOD SET_LRPROCESSCTRLINTVALUE
VAR_INPUT
	LRPROCESSCTRLINTVALUE : LREAL := 0.0;
END_VAR
END_METHOD

METHOD SET_LRPROCESSCTRLREDGAIN
VAR_INPUT
	LRPROCESSCTRLREDGAIN : LREAL := 0.0;
END_VAR
END_METHOD

METHOD SET_LRPROCESSCTRLREDRANGE
VAR_INPUT
	LRPROCESSCTRLREDRANGE : LREAL := 0.0;
END_VAR
END_METHOD

METHOD SET_RPROCESSCTRLDELAYTIME
VAR_INPUT
	RPROCESSCTRLDELAYTIME : REAL := 0.0;
END_VAR
END_METHOD

METHOD SET_RPROCESSCTRLRATEDTIME
VAR_INPUT
	RPROCESSCTRLRATEDTIME : REAL := 0.0;
END_VAR
END_METHOD

METHOD SET_XPICTRLLOADINTVALUE
VAR_INPUT
	XIN : BOOL := FALSE;
END_VAR
END_METHOD

METHOD SET_XPROCESSCTRLLOADINTVALUE
VAR_INPUT
	XPROCESSCTRLLOADINTVALUE : BOOL := FALSE;
END_VAR
END_METHOD

METHOD CALL_S000_CYCLIC
END_METHOD

METHOD CALL_S002_STANDBY
END_METHOD

METHOD CALL_S020_SYNCLINEVEL
END_METHOD

METHOD CALL_S050_DANCERTRL
END_METHOD

METHOD CALL_S999_ERROR
END_METHOD

METHOD CALL_T000_ALLSTATES
END_METHOD

METHOD CALL_T020_SYNCLINEVEL
END_METHOD

METHOD CALL_T050_DANCERTRL
END_METHOD

(* ---- L_TW2P_TM_WINDERDANCERCTRLSTATE.pou ---- *)
FUNCTION_BLOCK L_TW2P_TM_WINDERDANCERCTRLSTATE EXTENDS L_TW2P_TM_WinderDancerCtrlBase
VAR
	LRSETMINERTIAOUT : LREAL;
	LRIDENTMINERTIA : LREAL;
	LRSETSPDCTRLGAINADAPTOUT : LREAL;
	XDECOUPLINGACCCOMP : BOOL;
	LRACCTORQUE : LREAL;
	LRACTACCTORQUE : LREAL;
	XACCCMPSACTIVE_INT : BOOL;
	EDANCERCTRLSTOPMODE_OLD : L_TW2P_DancerCtrlStopMode;
	WSTEPPER_DANCERCTRLSTOPMODE : WORD;
	LRTIME : LREAL;
	LRDIST : LREAL;
	LRDISTTOTARGET : LREAL;
	LRRELDIST : LREAL;
	LRSTOREACTPOS : LREAL;
	LRPOS_DIST_INT : LREAL;
	LRTARGETPOSITION : LREAL;
	LRVEL_INT : LREAL;
	LRMAXMINERTIA : LREAL;
	XDONEFROMIDENTMINERTIA : BOOL;
	XIDENTMINERTIASPEELIMITS : BOOL;
	XEXECUTEIDENTDIAM_OLD : BOOL;
	WIDENTDIAMCALCCYCLES : WORD;
	XIDENTDIAMETERBUSY_INT : BOOL;
	XIDENTDIAMETERDONE_INT : BOOL;
	XIDENTDIAM_LOADDIAM : BOOL;
	LRIDENTDIAM_SETDIAMETER : LREAL;
	XERROR_IDENTDIAMMAXDANCERPOS : BOOL;
	XERROR_ACTDANPOSBIGGERMAXDANPOS : BOOL;
	XERRORFOLLOWINGERRORSWITCHTOPOSCTRLDRIVE : BOOL;
	XERROR_IDENTIFICATIONDIAMETERFAILED : BOOL;
	XERROR_INVALIDDANCERMATERIALLENGTH : BOOL;
	XWARNING_AXISNOTHOMEDSTOPMODEMOVEABS : BOOL;
	XWARNING_INVALIDDANCERMATERIALLENGTH : BOOL;
	XWARNING_IDENTIFICATIONDIAMETERFAILED : BOOL;
	XWARNING_INVALIDLOADDIAM : BOOL;
	XWARNING_INVALIDIDENTMAXDANCERPOS : BOOL;
	XWARNING_ACTDANCERPOSBIGGERMAXDANCERPOS : BOOL;
	L_MB1P_ACCCOMP1 : L_TB1P_AccComp;
	L_MB1P_IDENTMINERTIA1 : L_TB1P_IdentMInertia;
	L_MB1P_CURVESPEEDCTRLGAIN : L_USPP_Curve;
	FB_WINDERIDENTDIAMETER : L_TW2P_WinderIdentDiameter;
	FB_SETSPEEDCTRLADAPTVAL1 : L_MC1P_SetSpeedCtrlAdaptValue;
	ICTNSETSPEEDCTRLADAPTDISABLE : INT := 0;
END_VAR
END_FUNCTION_BLOCK

METHOD CALL_CTRLREQACTIVE : BOOL
END_METHOD

METHOD CALL_ERRORHANDLER
END_METHOD

METHOD CALL_FBMETHODS_WND
END_METHOD

METHOD CALL_FB_ACCCOMP : LREAL
END_METHOD

METHOD CALL_FB_CURVESPEEDCTRLGAIN
END_METHOD

METHOD CALL_FB_PROCESSCONTROLLER
END_METHOD

METHOD CALL_FB_SETSPEEDCTRLADAPTVALUE
END_METHOD

METHOD CALL_FB_WINDERIDENTDIAMETER
END_METHOD

METHOD CALL_FB_WNDCALCDIAMETER_INPUT
END_METHOD

METHOD CALL_FIRSTCYCLE
END_METHOD

METHOD CALL_INITROUTINE
END_METHOD

METHOD CALL_LIMITEDINPUT
END_METHOD

METHOD CALL_OUTPUT
END_METHOD

METHOD CALL_OUTPUT_SF
END_METHOD

METHOD CALL_REQUESTS_EXT
END_METHOD

METHOD CALL_RESETCOMMANDS
END_METHOD

METHOD CALL_RESETIDENTFBS
END_METHOD

METHOD CALL_RESETOUTPUT
END_METHOD

METHOD CALL_RESETWARNINGS
END_METHOD

METHOD CALL_SETSPEEDPOINT
END_METHOD

METHOD CALL_SETTORQUE
END_METHOD

METHOD CALL_STATEMACHINE
END_METHOD

METHOD CALL_WNDIDENTMINERTIA
END_METHOD

METHOD CALL_WNDTENSIONCURVE_INPUT
END_METHOD

METHOD CALL_ABC_INPUT
END_METHOD

METHOD CALL_ABC_INPUT_PROFILEPARAMETER
END_METHOD

METHOD GET_LRACTACCTRQ : LREAL
END_METHOD

METHOD CALL_S000_CYCLIC
END_METHOD

METHOD CALL_S002_STANDBY
END_METHOD

METHOD CALL_S014_MOVEABS
END_METHOD

METHOD CALL_S015_LINEJOGGING
END_METHOD

METHOD CALL_S015_MOVEREL
END_METHOD

METHOD CALL_S020_SYNCLINEVEL
END_METHOD

METHOD CALL_S040_IDENTMINERTIA
END_METHOD

METHOD CALL_S050_DANCERTRL
END_METHOD

METHOD CALL_S081_IDENTDIAMETER
END_METHOD

METHOD CALL_S996_STOP
END_METHOD

METHOD CALL_S999_ERROR
END_METHOD

METHOD CALL_T000_ALLSTATES
END_METHOD

METHOD CALL_T050_DANCERTRL
END_METHOD

(* ---- L_TW2P_TM_WINDERTENSIONCTRLBASE.pou ---- *)
FUNCTION_BLOCK L_TW2P_TM_WINDERTENSIONCTRLBASE EXTENDS L_TW2P_TM_Winder
VAR_OUTPUT
	PPAR : POINTER TO L_TW2P_scPar_TM_WinderTensionCtrlState := ADR(scPar_int);
	PSF : POINTER TO L_TW2P_scSF_TM_WinderTensionCtrlState;
	PAP : POINTER TO L_TW2P_scAP_TM_WinderTensionCtrlState;
END_VAR
VAR
	PINPUTWINDERTENS : POINTER TO L_TW2P_WinderTensionCtrlStateIn;
	POUTPUTWINDERTENS : POINTER TO L_TW2P_WinderTensionCtrlStateOut;
	TM_WINDERDANCERCTRLBASECONFIG : L_TB2P_ModuleHandlerConfig;
	XCONSTANTTENSION : BOOL;
	XWNDSPDLIMIT : BOOL;
	LRSETMINERTIAOUT : LREAL;
	XTENSINTARGET : BOOL;
	LRACTTENSIN_INT : LREAL := 0;
	LRFILTACTTENSIN : LREAL;
	XPICONTROLACTIVE_INT : BOOL;
	SCPAR_INT : L_TW2P_scPar_TM_WinderTensionCtrlState;
	WTENSRAMPLOADSTARTVALUEMODE : WORD;
	LRSETTENSSCALED : LREAL;
	LRPROCESSCTRLREDOUT : LREAL;
	LRSETPOINTTENSION : LREAL;
	LRSETTENSIONTORQUE : LREAL;
	LRSETFRICTIONTORQUE : LREAL;
	LRACTFRICTIONTORQUE : LREAL;
	LRACCTORQUE : LREAL;
	LRACTACCTORQUE : LREAL;
	LRSETLINEVELOFFSET : LREAL;
	LRSETTRQPOINT : LREAL;
	LRCALCWNDSPEEDUPPERLIMIT : LREAL;
	LRCALCWNDSPEEDLOWERLIMIT : LREAL;
	XACCCMPSACTIVE_INT : BOOL;
	XDECOUPLINGACCCOMP : BOOL;
	XDECOUPLINGFRICTIONCOMP : BOOL;
	XDECOUPLINGTENSION : BOOL;
	LRMAXMINERTIA : LREAL;
	ETENSCTRLMODE_LOCK : L_TW2P_WinderTensionControlMode := L_TW2P_WinderTensionControlMode.TorqueBased;
	XWNDSPDLIMIT_OLD : BOOL;
	ICNTSPDLIMIT : INT;
	ISPDHYST : INT := 3;
	XACTTENSINTARGET_INT : BOOL;
	LRTENSINWINDOW_INT : LREAL;
	L_MB1P_ACCCOMP1 : L_TB1P_AccComp;
	L_D94A_FILTERREELSPEED : L_USPP_PT1Filter;
	L_D94A_FILTERREELSPEEDFRICTIONCOMP : L_USPP_PT1Filter;
END_VAR
END_FUNCTION_BLOCK

METHOD CALL_ALLOCPOINTADR
END_METHOD

METHOD CALL_CTRLREQACTIVE : BOOL
END_METHOD

METHOD CALL_FBMETHODS_WND
END_METHOD

METHOD CALL_FB_ACCCOMP : LREAL
END_METHOD

METHOD CALL_FB_ACCCOMP_INPUT : LREAL
END_METHOD

METHOD CALL_FB_RAMPGENERATOR_INPUT
END_METHOD

METHOD CALL_FB_WNDCALCDIAMETER_INPUT
END_METHOD

METHOD CALL_FILTERREELSPEED
END_METHOD

METHOD CALL_FIRSTCYCLE
END_METHOD

METHOD CALL_INTERNALCTRL
END_METHOD

METHOD CALL_OUTPUT
END_METHOD

METHOD CALL_OUTPUT_SF
END_METHOD

METHOD CALL_REQUESTS_EXT
END_METHOD

METHOD CALL_RESETCOMMANDS
END_METHOD

METHOD CALL_RESETOUTPUT
END_METHOD

METHOD CALL_SDRAMPGENERATOR_INPUT
END_METHOD

METHOD CALL_SETTORQUE
END_METHOD

METHOD CALL_SPEEDLIMIT
END_METHOD

METHOD CALL_STATEMACHINE
END_METHOD

METHOD CALL_WNDFRICTIONCOMPENSATION
END_METHOD

METHOD GET_LRACTACCTRQ : LREAL
END_METHOD

METHOD GET_LRACTFRICTRQ : LREAL
END_METHOD

METHOD GET_LRACTTENSTRQ : LREAL
END_METHOD

METHOD GET_LRRAMPGENOUT : LREAL
END_METHOD

METHOD GET_LRSPEEDLOWERLIMIT : LREAL
END_METHOD

METHOD GET_LRSPEEDUPPERLIMIT : LREAL
END_METHOD

METHOD GET_LRTENSCTRLOUT : LREAL
END_METHOD

METHOD GET_LRTENSCURVEOUT : LREAL
END_METHOD

METHOD CALL_S000_CYCLIC
END_METHOD

METHOD CALL_S015_LINEJOGGING
END_METHOD

METHOD CALL_S020_SYNCLINEVEL
END_METHOD

METHOD CALL_S050_1_WNDFRICTIONCOMPENSATION
END_METHOD

METHOD CALL_S050_TENSIONCTRL
END_METHOD

METHOD CALL_T000_ALLSTATES
END_METHOD

METHOD CALL_T020_SYNCLINEVEL
END_METHOD

METHOD CALL_T050_TENSIONCTRL
END_METHOD

(* ---- L_TW2P_TM_WINDERTENSIONCTRLSTATE.pou ---- *)
FUNCTION_BLOCK L_TW2P_TM_WINDERTENSIONCTRLSTATE EXTENDS L_TW2P_TM_WinderTensionCtrlBase
VAR_IN_OUT
	ALRFRICTIONCURVE1 : ARRAY [1..66] OF LREAL;
	ALRFRICTIONCURVE2 : ARRAY [1..66] OF LREAL;
	ALRFRICTIONCURVE3 : ARRAY [1..66] OF LREAL;
	ALRFRICTIONCURVE4 : ARRAY [1..66] OF LREAL;
END_VAR
VAR
	LRIDENTMINERTIA : LREAL;
	LRSETSPDCTRLGAINADAPTOUT : LREAL;
	XRESETPICTRL_OLD : BOOL;
	XRESETICTRL_OLD : BOOL;
	LRTENSCTRLRESETTIME_STORE : LREAL;
	LRDEVIATION_STORE : LREAL;
	LRPROCESSCTRLREDOUTVEL : LREAL;
	LRSETREELSPEEDFRWCTRL : LREAL;
	LRTENSCTRLLIMITNEG_INT : LREAL;
	LRTENSCTRLLIMITPOS_INT : LREAL;
	WSTEPPER_TENSCTRLSTOPMODE : WORD;
	ESTOPMODE_OLD : L_TW2P_TensionCtrlStopMode;
	LRRELDIST : LREAL;
	LRSTOREACTPOS : LREAL;
	LRDISTTOTARGET : LREAL;
	LRVEL_INT : LREAL;
	LRTARGETPOSITION : LREAL;
	LRDIST : LREAL;
	LRTIME : LREAL;
	LRVELOCITY_OLD : LREAL;
	XIDENTMINERTIASPEELIMITS : BOOL;
	XDONEFROMIDENTMINERTIA : BOOL;
	XPIDENABLE_INT : BOOL;
	XPIDRESET_INT : BOOL;
	XPIDLOADACTVLAUE_INT : BOOL;
	XPIDLRESETICTRLACTIVE_INT : BOOL;
	XPIDLRESETPICTRLACTIVE_INT : BOOL;
	LRTENSPICTRLOUT : LREAL;
	LRHYSTERISWIDTH : LREAL;
	XERRORFOLLOWINGERRORSWITCHTOPOSCTRLDRIVE : BOOL;
	L_MB1P_RAMPGENERATORRESETICTRL : L_MC1P_RampGenerator;
	L_MB1P_RAMPGENERATORRESETPICTRL : L_MC1P_RampGenerator;
	XRAMPGENSETVALUEFORPICTRLACTIVE : BOOL;
	WRESETPICTRL_STEPPER : WORD;
	L_MB1P_PROCESSCONTROLLER1 : L_CT1P_ProcessController;
	L_MB1P_FRICTIONCOMPENSATION1 : L_TB1P_FrictionCompensation;
	L_D94A_FILTERTENSIN : L_USPP_PT1Filter;
	L_MB1P_IDENTMINERTIA1 : L_TB1P_IdentMInertia;
	L_MB1P_CURVESPEEDCTRLGAIN : L_USPP_Curve;
	FB_SETSPEEDCTRLADAPTVAL1 : L_MC1P_SetSpeedCtrlAdaptValue;
	ICTNSETSPEEDCTRLADAPTDISABLE : INT := 1;
END_VAR
END_FUNCTION_BLOCK

METHOD CALL_CTRLREQACTIVE : BOOL
END_METHOD

METHOD CALL_ERRORHANDLER
END_METHOD

METHOD CALL_FBMETHODS_WND
END_METHOD

METHOD CALL_FB_CURVESPEEDCTRLGAIN
END_METHOD

METHOD CALL_FB_CURVESPEEDCTRLGAIN_INPUT
END_METHOD

METHOD CALL_FB_PROCESSCONTROLLER
END_METHOD

METHOD CALL_FB_PROCESSCONTROLLER_INPUT
END_METHOD

METHOD CALL_FB_RAMGENERATORRESETPICTRL
END_METHOD

METHOD CALL_FB_RAMPGENERATORRESETICTRL
END_METHOD

METHOD CALL_FB_RAMPGENERATORRESETICTRL_INPUT
END_METHOD

METHOD CALL_FB_RAMPGENERATORRESETPICTRL_INPUT
END_METHOD

METHOD CALL_FB_SETSPEEDCTRLADAPTVALUE
END_METHOD

METHOD CALL_FB_SETSPEEDCTRLADAPTVALUE_INPUT
END_METHOD

METHOD CALL_FILTERTENSIN
END_METHOD

METHOD CALL_FIRSTCYCLE
END_METHOD

METHOD CALL_INITROUTINE
END_METHOD

METHOD CALL_INTERNALCTRL
END_METHOD

METHOD CALL_LIMITEDINPUT
END_METHOD

METHOD CALL_OUTPUT
END_METHOD

METHOD CALL_OUTPUT_SF
END_METHOD

METHOD CALL_REQUESTS_EXT
END_METHOD

METHOD CALL_RESETCOMMANDS
END_METHOD

METHOD CALL_RESETIDENTFBS
END_METHOD

METHOD CALL_RESETOUTPUT
END_METHOD

METHOD CALL_SETSPEEDPOINT
END_METHOD

METHOD CALL_SETTORQUE
END_METHOD

METHOD CALL_SETWINDERID
END_METHOD

METHOD CALL_STATEMACHINE
END_METHOD

METHOD CALL_WNDFRICTIONCOMPENSATION
END_METHOD

METHOD CALL_WNDIDENTMINERTIA
END_METHOD

METHOD CALL_WNDTENSIONCURVE_INPUT
END_METHOD

METHOD CALL_ABC_INPUT
END_METHOD

METHOD CALL_ABC_INPUT_PROFILEPARAMETER
END_METHOD

METHOD SET_ALRPROCESSCTRLXVALUES
VAR_INPUT
	ALRPROCESSCTRLXVALUES : ARRAY [1..5] OF LREAL;
END_VAR
END_METHOD

METHOD SET_ALRPROCESSCTRLYVALUES
VAR_INPUT
	ALRPROCESSCTRLYVALUES : ARRAY [1..5] OF LREAL;
END_VAR
END_METHOD

METHOD SET_LRPICTRLINTVALUE
VAR_INPUT
	LRIN : LREAL := 0;
END_VAR
END_METHOD

METHOD SET_LRPROCESSCTRLACC
VAR_INPUT
	LRPROCESSCTRLACC : LREAL := 0.0;
END_VAR
END_METHOD

METHOD SET_LRPROCESSCTRLDEC
VAR_INPUT
	LRPROCESSCTRLDEC : LREAL := 0.0;
END_VAR
END_METHOD

METHOD SET_LRPROCESSCTRLGAINADAPT
VAR_INPUT
	LRPROCESSCTRLGAINADAPT : LREAL := 1;
END_VAR
END_METHOD

METHOD SET_LRPROCESSCTRLINTVALUE
VAR_INPUT
	LRPROCESSCTRLINTVALUE : LREAL := 0.0;
END_VAR
END_METHOD

METHOD SET_LRPROCESSCTRLREDGAIN
VAR_INPUT
	LRPROCESSCTRLREDGAIN : LREAL := 0.0;
END_VAR
END_METHOD

METHOD SET_LRPROCESSCTRLREDRANGE
VAR_INPUT
	LRPROCESSCTRLREDRANGE : LREAL := 0.0;
END_VAR
END_METHOD

METHOD SET_RPROCESSCTRLDELAYTIME
VAR_INPUT
	RPROCESSCTRLDELAYTIME : REAL := 0.0;
END_VAR
END_METHOD

METHOD SET_RPROCESSCTRLRATEDTIME
VAR_INPUT
	RPROCESSCTRLRATEDTIME : REAL := 0.0;
END_VAR
END_METHOD

METHOD SET_XPICTRLLOADINTVALUE
VAR_INPUT
	XIN : BOOL := FALSE;
END_VAR
END_METHOD

METHOD SET_XPROCESSCTRLLOADINTVALUE
VAR_INPUT
	XPROCESSCTRLLOADINTVALUE : BOOL := FALSE;
END_VAR
END_METHOD

METHOD CALL_S000_CYCLIC
END_METHOD

METHOD CALL_S002_STANDBY
END_METHOD

METHOD CALL_S014_MOVEABS
END_METHOD

METHOD CALL_S015_MOVEREL
END_METHOD

METHOD CALL_S030_IDENTFRICTION
END_METHOD

METHOD CALL_S040_IDENTMINERTIA
END_METHOD

METHOD CALL_S050_1_WNDFRICTIONCOMPENSATION
END_METHOD

METHOD CALL_S050_TENSIONCTRL
END_METHOD

METHOD CALL_S996_STOP
END_METHOD

METHOD CALL_S999_ERROR
END_METHOD

METHOD CALL_T000_ALLSTATES
END_METHOD

METHOD CALL_T020_SYNCLINEVEL
END_METHOD

METHOD CALL_T050_TENSIONCTRL
END_METHOD

(* ---- L_TW2P_WINDER.pou ---- *)
FUNCTION_BLOCK L_TW2P_WINDER EXTENDS L_TB2P_TechModuleBase
END_FUNCTION_BLOCK

METHOD CALL_SMC_READPARAMETEREXT
VAR_INPUT
	XENABLE : BOOL;
	WCODENUMBER : WORD;
	BYSUBCODE : BYTE;
END_VAR
VAR_OUTPUT
	XVALID : BOOL;
	XBUSY : BOOL;
	XERROR : BOOL;
	WERRORID : WORD;
	DWVALUE : DWORD;
END_VAR
END_METHOD

METHOD CALL_WRITEPARAMETEREXT
VAR_INPUT
	XEXECUTE : BOOL;
	WCODENUMBER : WORD;
	BYSUBCODE : BYTE;
	BYLENGTH : BYTE;
	DNVALUE : DINT;
END_VAR
VAR_OUTPUT
	XDONE : BOOL;
	XBUSY : BOOL;
	XERROR : BOOL;
	WERRORID : WORD;
END_VAR
END_METHOD

METHOD CALL_WRITEPARAMETEREXT2
VAR_INPUT
	XEXECUTE : BOOL;
	WCODENUMBER : WORD;
	BYSUBCODE : BYTE;
	BYLENGTH : BYTE;
	DNVALUE : DINT;
END_VAR
VAR_OUTPUT
	XDONE : BOOL;
	XBUSY : BOOL;
	XERROR : BOOL;
	WERRORID : WORD;
END_VAR
END_METHOD

METHOD GET_ESTATE : L_TB2P_States
END_METHOD

METHOD GET_ETMSTATE : L_TB2P_States
END_METHOD

METHOD GET_FSCALEFACTOR : LREAL
END_METHOD

METHOD GET_LRACTMOTORTORQUE : LREAL
END_METHOD

METHOD GET_LRCALCDIAMDIST : LREAL
END_METHOD

METHOD GET_LRFEEDCONSTANT : LREAL
END_METHOD

METHOD GET_LRLOWERSPEEDLIMIT : LREAL
END_METHOD

METHOD GET_LRMOTORTORQUEREF : LREAL
END_METHOD

METHOD GET_LRREELSPEEDREF : LREAL
END_METHOD

METHOD GET_LRSETMOTORTORQUE : LREAL
END_METHOD

METHOD GET_LRSETSPEEDCTRLGAINADAPT : LREAL
END_METHOD

METHOD GET_LRSETTOTALTORQUE : LREAL
END_METHOD

METHOD GET_LRTASKCYCLE : LREAL
END_METHOD

METHOD GET_LRUPPERSPEEDLIMIT : LREAL
END_METHOD

METHOD GET_LRVARMINERTIASCALED : LREAL
END_METHOD

METHOD GET_LRWINDERTORQUEREF : LREAL
END_METHOD

METHOD GET_WCHECKAXISTYP : WORD
END_METHOD

METHOD GET_XCOMMUNICATION : BOOL
END_METHOD

METHOD GET_XDIAMWEBBREAKENABLE : BOOL
VAR_OUTPUT
	XUNIDIRECT : BOOL;
	XUNWINDACTIVE : BOOL;
END_VAR
END_METHOD

METHOD RESET_SYSTEMFAULT
END_METHOD

METHOD SET_SYSTEMFAULT
VAR_INPUT
	IN : L_IE1P_Error;
END_VAR
END_METHOD

METHOD SET_WNDAXISEXTENSION_READY
END_METHOD

METHOD SET_ESTATE
VAR_INPUT
	IN : L_TB2P_States;
END_VAR
END_METHOD

METHOD SET_LRFEEDCONSTANT
VAR_INPUT
	LRIN : LREAL := 0;
END_VAR
END_METHOD

METHOD SET_LRREFERENCEMOTORTORQUE
VAR_INPUT
	LRIN : LREAL := 0;
END_VAR
END_METHOD

METHOD SET_LRREFERENCEREELSPEED
VAR_INPUT
	LRIN : LREAL := 0;
END_VAR
END_METHOD

METHOD SET_LRSPEEDOFFSET
VAR_INPUT
	LRIN : LREAL := 0;
END_VAR
END_METHOD

METHOD SET_LRTORQUEOFFSET
VAR_INPUT
	LRIN : LREAL := 0;
END_VAR
END_METHOD

METHOD SET_XSPEEDLIMITENABLEDEXT
VAR_INPUT
	XIN : BOOL := TRUE;
END_VAR
END_METHOD

METHOD SET_XWEBBREAK
VAR_INPUT
	XIN : BOOL := FALSE;
END_VAR
END_METHOD

(* ---- L_TW2P_WINDERDANCERCTRLSTATE.pou ---- *)
FUNCTION_BLOCK L_TW2P_WINDERDANCERCTRLSTATE EXTENDS L_TW2P_Winder
VAR_INPUT
	XENABLE : BOOL;
	XENABLEOPERATION : BOOL;
	XRESETERROR : BOOL;
	XQSPAPPLICATION : BOOL;
	XABORT : BOOL;
	XJOGPOS : BOOL;
	XJOGNEG : BOOL;
	XHOMEEXECUTE : BOOL;
	LROVERRIDE : LREAL := 1;
	SCCTRLBASICMOTION : L_TB2P_scCtrlBasicMotion;
	SCPAR : L_TW2P_scPar_WinderDancerCtrlState;
	SCACCESSPOINTS : L_TW2P_scAP_WinderDancerCtrlState;
	XMATERIALFEEDING : BOOL;
	XWINDINGDIRECTION : BOOL;
	XJOGLINEPOS : BOOL;
	XJOGLINENEG : BOOL;
	LRSETLINEVEL : LREAL;
	LRSETLINEVELDIAMCALC : LREAL;
	XLOADDIAM : BOOL;
	LRLOADDIAM : LREAL;
	XHOLDDIAM : BOOL;
	XDIAMCALCREDUCED : BOOL;
	XWEBBREAKMONIT : BOOL;
	XSYNCIN : BOOL;
	XTEACHUPPERPOS : BOOL;
	XTEACHLOWERPOS : BOOL;
	LRACTDANCERPOSIN : LREAL;
	XDANCERCTRL : BOOL;
	LRSETDANCERPOSSCALED : LREAL;
	LRCTRLINFLUENCESCALED : LREAL;
	XRESETICTRL : BOOL;
	XACCCMPS : BOOL;
	LRMINERTIAADAPT : LREAL := 1;
	XEXECUTEIDENTMINERTIA : BOOL;
	XEXECUTEIDENTDIAM : BOOL;
	XADAPTSPDCTRLGAIN : BOOL;
	LRADAPTSPDCTRLGAINFACTOR : LREAL := 1;
	XTENSCURVE : BOOL;
	LRSETTENS : LREAL;
	XSETMATERIALCOUNTER : BOOL;
	MATERIALCOUNTERVALUES : L_MC1P_IAXIS_REF_MASTERVALUES;
END_VAR
VAR_OUTPUT
	XREADYFOROPERATION : BOOL;
	XOPERATIONENABLED : BOOL;
	XREADYFORMOTION : BOOL;
	XERROR : BOOL;
	XWARNING : BOOL;
	EERRORID : L_IE1P_Error;
	XSTOACTIVE : BOOL;
	XQSPACTIVE : BOOL;
	XABORTBUSY : BOOL;
	XABORTDONE : BOOL;
	XJOGGINGBUSY : BOOL;
	XHOMINGBUSY : BOOL;
	XHOMINGDONE : BOOL;
	XISHOMED : BOOL;
	ETMSTATE : L_TB2P_States := L_TB2P_States.DISABLED;
	SCSTATUSBASICMOTION : L_TB2P_scStatusBasicMotion;
	LRACTVEL : LREAL;
	LRSETVELOUT : LREAL;
	LRACTPOS : LREAL;
	LRSETPOSOUT : LREAL;
	LRACTFOLLOWINGERROR : LREAL;
	SCSIGNALFLOW : L_TW2P_scSF_WinderDancerCtrlState;
	XHOLDDIAMACTIVE : BOOL;
	XDIAMMAX : BOOL;
	XDIAMMIN : BOOL;
	LRSETDIAMOUT : LREAL;
	XWEBBREAK : BOOL;
	XSYNCHRONISED : BOOL;
	XACCDECSYNC : BOOL;
	XWINDINGBUSY : BOOL;
	XUNWIND : BOOL;
	LRACTDANCERPOSSCALED : LREAL;
	XDANCERREACHEDSETPOS : BOOL;
	XDANCERMAXPOS : BOOL;
	XDANCERMINPOS : BOOL;
	LRSETMINERTIAOUT : LREAL;
	XIDENTBUSY : BOOL;
	XIDENTDONE : BOOL;
	LRIDENTMINERTIA : LREAL;
	LRSETSPDCTRLGAINADAPTOUT : LREAL;
	LRSETTENSCURVEOUT : LREAL;
	LRMATERIALCOUNTER : LREAL;
	LRLIMITLINEVEL : LREAL;
	XVELOCITYMASTERBUSY : BOOL;
	LRSETLINEVELOUT : LREAL;
	XLINESTOP : BOOL;
END_VAR
VAR_IN_OUT
	AXIS : AXIS_REF;
	PERSISTENTVAR : L_TW2P_PersistentVarWinder;
END_VAR
VAR
	TM_INT : L_TW2P_TM_WinderDancerCtrlState := STRUCT(ModuleHandler := ModuleHandler);
	_UICALLMFUNIDXINPUT : UINT := 1;
	_UICALLMFUNIDXOUTPUT : UINT := 1;
	_ASCINPUT : ARRAY [1.._MCCall.c_BufferDepthInput] OF L_TW2P_WinderDancerCtrlStateIn;
	_ASCOUTPUT : ARRAY [1.._MCCall.c_BufferDepthOutput] OF L_TW2P_WinderDancerCtrlStateOut;
	_ASCPARCORE : ARRAY [1.._MCCall.c_BufferDepthInput] OF L_TW2P_scPar_WinderDancerCtrlState;
	_MCCALL : L_UM1P_MCCall;
	_ASCACCESSPOINTSCORE : ARRAY [1.._MCCall.c_BufferDepthInput] OF L_TW2P_scAP_WinderDancerCtrlState;
	_ASCSIGNALFLOWCORE : ARRAY [1.._MCCall.c_BufferDepthOutput] OF L_TW2P_scSF_WinderDancerCtrlState;
	SCPAR_INT : L_TW2P_scPar_WinderDancerCtrlState;
	_SCINPUTVISU : L_TW2P_WinderDancerCtrlStateIn;
	_PSCINPUTVISU : POINTER TO L_TW2P_WinderDancerCtrlStateIn := ADR(_scInputVisu);
	_PSCOUTPUTVISU : POINTER TO L_TW2P_WinderDancerCtrlStateOut := ADR(_ascOutput[1]);
	_PSCPARVISU : POINTER TO L_TW2P_scPar_WinderDancerCtrlState := ADR(scPar_int);
	ITFITECHMODULEINTERNAL : L_TB2P_ITechModuleInternal;
	LRJERKDEC : LREAL;
	LRJOGGINGJERKDEC : LREAL;
	REMAININGTIMEOFPROFILE : LREAL;
	REMAININGTIMEOFPROFILEAVAILABLE : BOOL;
END_VAR
END_FUNCTION_BLOCK

METHOD CALL_COUPLINGREELSPEEDLIMIT
END_METHOD

METHOD CALL_DECOUPLINGREELSPEEDLIMIT
END_METHOD

METHOD CALL_RESTDANCERTEACHPOS
END_METHOD

METHOD GET_ESTATE : L_TB2P_States
END_METHOD

METHOD GET_ETMSTATE : L_TB2P_States
END_METHOD

METHOD GET_LRACTACCTRQ : LREAL
END_METHOD

METHOD GET_LRACTDANCERCTRLOUT : LREAL
END_METHOD

METHOD GET_LRACTDANCERLINEVELCOMP : LREAL
END_METHOD

METHOD GET_LRACTDANCERVEL : LREAL
END_METHOD

METHOD GET_LRACTMOTORTORQUE : LREAL
END_METHOD

METHOD GET_LRCALCDIAMDIST : LREAL
END_METHOD

METHOD GET_LRCALCDIAMLINESPEED : LREAL
END_METHOD

METHOD GET_LRCALCDIAMREELSPEED : LREAL
END_METHOD

METHOD GET_LRFEEDCONSTANT : LREAL
END_METHOD

METHOD GET_LRLOWERSPEEDLIMIT : LREAL
END_METHOD

METHOD GET_LRMOTORTORQUEREF : LREAL
END_METHOD

METHOD GET_LRREELSPEEDREF : LREAL
END_METHOD

METHOD GET_LRSETMOTORTORQUE : LREAL
END_METHOD

METHOD GET_LRSETSPEEDCTRLGAINADAPT : LREAL
END_METHOD

METHOD GET_LRSETTOTALTORQUE : LREAL
END_METHOD

METHOD GET_LRSPEEDFORWARDCTRL : LREAL
END_METHOD

METHOD GET_LRSPEEDSETPOINT : LREAL
END_METHOD

METHOD GET_LRTASKCYCLE : LREAL
END_METHOD

METHOD GET_LRUPPERSPEEDLIMIT : LREAL
END_METHOD

METHOD GET_LRVARMINERTIASCALED : LREAL
END_METHOD

METHOD GET_LRVELSETPOINT : LREAL
END_METHOD

METHOD GET_LRWINDERTORQUEREF : LREAL
END_METHOD

METHOD GET_XCOMMUNICATION : BOOL
END_METHOD

METHOD GET_XDIAMWEBBREAKENABLE : BOOL
VAR_OUTPUT
	XUNIDIRECT : BOOL;
	XUNWINDACTIVE : BOOL;
END_VAR
END_METHOD

METHOD GET_XLOWERPOSTEACHED : BOOL
VAR_OUTPUT
	LRTEACHPOSLOWERLIMIT : LREAL;
END_VAR
END_METHOD

METHOD GET_XUPPERPOSTEACHED : BOOL
VAR_OUTPUT
	LRTEACHPOSUPPERLIMIT : LREAL;
END_VAR
END_METHOD

METHOD LOAD_LRDANCERLOWERLIMIT
VAR_INPUT
	LRIN : LREAL := 0;
END_VAR
END_METHOD

METHOD LOAD_LRDANCERUPPERLIMIT
VAR_INPUT
	LRIN : LREAL := 0;
END_VAR
END_METHOD

METHOD SET_ALRPROCESSCTRLXVALUES
VAR_INPUT
	ALRPROCESSCTRLXVALUES : ARRAY [1..5] OF LREAL;
END_VAR
END_METHOD

METHOD SET_ALRPROCESSCTRLYVALUES
VAR_INPUT
	ALRPROCESSCTRLYVALUES : ARRAY [1..5] OF LREAL;
END_VAR
END_METHOD

METHOD SET_ESTATE
VAR_INPUT
	IN : L_TB2P_States;
END_VAR
END_METHOD

METHOD SET_LRFEEDCONSTANT
VAR_INPUT
	LRIN : LREAL := 0;
END_VAR
END_METHOD

METHOD SET_LRPICTRLINTVALUE
VAR_INPUT
	LRIN : LREAL := 0;
END_VAR
END_METHOD

METHOD SET_LRPROCESSCTRLACC
VAR_INPUT
	LRPROCESSCTRLACC : LREAL := 0.0;
END_VAR
END_METHOD

METHOD SET_LRPROCESSCTRLDEC
VAR_INPUT
	LRPROCESSCTRLDEC : LREAL := 0.0;
END_VAR
END_METHOD

METHOD SET_LRPROCESSCTRLGAINADAPT
VAR_INPUT
	LRPROCESSCTRLGAINADAPT : LREAL := 1;
END_VAR
END_METHOD

METHOD SET_LRPROCESSCTRLINTVALUE
VAR_INPUT
	LRPROCESSCTRLINTVALUE : LREAL := 0.0;
END_VAR
END_METHOD

METHOD SET_LRPROCESSCTRLREDGAIN
VAR_INPUT
	LRPROCESSCTRLREDGAIN : LREAL := 0.0;
END_VAR
END_METHOD

METHOD SET_LRPROCESSCTRLREDRANGE
VAR_INPUT
	LRPROCESSCTRLREDRANGE : LREAL := 0.0;
END_VAR
END_METHOD

METHOD SET_LRREFERENCEMOTORTORQUE
VAR_INPUT
	LRIN : LREAL := 0;
END_VAR
END_METHOD

METHOD SET_LRREFERENCEREELSPEED
VAR_INPUT
	LRIN : LREAL := 0;
END_VAR
END_METHOD

METHOD SET_LRSPEEDOFFSET
VAR_INPUT
	LRIN : LREAL := 0;
END_VAR
END_METHOD

METHOD SET_LRTORQUEOFFSET
VAR_INPUT
	LRIN : LREAL := 0;
END_VAR
END_METHOD

METHOD SET_RPROCESSCTRLDELAYTIME
VAR_INPUT
	RPROCESSCTRLDELAYTIME : REAL := 0.0;
END_VAR
END_METHOD

METHOD SET_RPROCESSCTRLRATEDTIME
VAR_INPUT
	RPROCESSCTRLRATEDTIME : REAL := 0.0;
END_VAR
END_METHOD

METHOD SET_XPICTRLLOADINTVALUE
VAR_INPUT
	XIN : BOOL := FALSE;
END_VAR
END_METHOD

METHOD SET_XPROCESSCTRLLOADINTVALUE
VAR_INPUT
	XPROCESSCTRLLOADINTVALUE : BOOL := FALSE;
END_VAR
END_METHOD

METHOD SET_XSPEEDLIMITENABLEDEXT
VAR_INPUT
	XIN : BOOL := TRUE;
END_VAR
END_METHOD

METHOD SET_XWEBBREAK
VAR_INPUT
	XIN : BOOL := FALSE;
END_VAR
END_METHOD

METHOD CALLFUNCTION
VAR_INPUT
	UIINPUTDATAIDX : UINT;
	UIOUTPUTDATAIDX : UINT;
END_VAR
END_METHOD

METHOD COPYINPUTS : BOOL
VAR_INPUT
	IDX : WORD;
END_VAR
END_METHOD

METHOD COPYOUTPUTS : BOOL
VAR_INPUT
	IDX : WORD;
END_VAR
END_METHOD

METHOD FUNCTIONWASCALLEDTWICE : BOOL
VAR_INPUT
	IDX : WORD;
END_VAR
END_METHOD

METHOD HANDLESTANDARDCALL : BOOL
END_METHOD

METHOD SYNCOUTPUTS
VAR_INPUT
	UICOPYOUTPUTFROMIDX : UINT;
	UICOPYOUTPUTTOIDX : UINT;
END_VAR
END_METHOD

METHOD CALL_INTERNALCTRL
END_METHOD

METHOD GET_PAP : POINTER TO L_TB2P_scAP_TM_MotionControl
END_METHOD

METHOD GET_PPAR : POINTER TO L_TB2P.L_TB2P_scPar_TM_MotionControl
END_METHOD

METHOD GET_PSF : POINTER TO L_TB2P_scSF_TM_MotionControl
END_METHOD

(* ---- L_TW2P_WINDERIDENTDIAMETER.pou ---- *)
FUNCTION_BLOCK L_TW2P_WINDERIDENTDIAMETER
VAR_INPUT
	XEXECUTE : BOOL;
	XABORT : BOOL;
	XDANCERMINPOS : BOOL;
	LRACTREELSPEEDIN : LREAL;
	LRACTDANCERPOSIN : LREAL;
	XLINEVELDIAMCALC : BOOL;
	LRSETLINEVELDIAMCALC : LREAL;
	LRMAXDANCERPOS : LREAL;
	LRDANCERMATERIALLENGTH : LREAL;
	LRMAXDIAM : LREAL;
	LRDIAMCALCDIST : LREAL;
	WIDENTDIAMCALCCYCLES : WORD := 1;
	LRTASKCYCLE : LREAL := 0.001;
	LRIDENTVEL : LREAL;
	LRIDENTACC : LREAL;
	LRIDENTDEC : LREAL;
	LRIDENTJERK : LREAL;
END_VAR
VAR_OUTPUT
	XERROR : BOOL;
	EERRORID : WORD;
	XBUSY : BOOL;
	XDONE : BOOL;
	XCOMMANDABORTED : BOOL;
	LRSETREELSPEEDOUT : LREAL;
	LRIDETDIAM : LREAL;
END_VAR
VAR
	WSTATE : WORD;
	LRTASKCYCLE_INT : LREAL := 0.001;
	LRMAXDIAM_INT : LREAL;
	LRREELSPEEDFAKTOR_INT : LREAL;
	LRMAXDANCERPOS_INT : LREAL;
	LRDANCERMATERIALLENGTH_INT : LREAL;
	XLINEVELDIAMCALC_INT : BOOL;
	LRREELSPEEDOUT_INT : LREAL;
	LRACTREELDIST_INT : LREAL;
	LRACTDIST_INT : LREAL;
	LRPROFGENDIST_INT : LREAL;
	LRSETDIST_INT : LREAL;
	LRSETDISTCALCDIAM_INT : LREAL;
	LRPROFGENSTARTPOSIDENTDIAM_INT : LREAL;
	LRPROFGENENDPOSIDENTDIAM_INT : LREAL;
	LRRAMPGENDECDIST : LREAL;
	XRAMPGENHALT : BOOL;
	XIDENTSTARTVALUESVALID : BOOL;
	XIDENTENDVALUESVALID : BOOL;
	LRDANCERPOSSTARTIDENT : LREAL;
	LRDANCERPOSENDIDENT : LREAL;
	LRLINEVELSTARTIDENT : LREAL;
	LRLINEVELENDIDENT : LREAL;
	LRLINEDIST : LREAL;
	LRWNDPOSSTARTIDENT : LREAL;
	LRWNDPOSENDIDENT : LREAL;
	LRIDETNWINDDIST : LREAL;
	XERROR_INVALIDMAXDIAM : BOOL;
	XERROR_INVALIDDANCERMATERIALLENGTH : BOOL;
	XERROR_ACTDANPOSBIGGERMAXDANPOS : BOOL;
	XERROR_ACTDANPOSBIGGERMAXDANPOS_TMP : BOOL;
	XEXECUTE_OLD : BOOL;
	XABORT_OLD : BOOL;
	FB_RAMPGENERATOR1 : L_MC1P_RampGenerator;
END_VAR
END_FUNCTION_BLOCK

METHOD CALL_ERRORHANDLER
END_METHOD

METHOD CALL_FBMETHODS
END_METHOD

METHOD CALL_FB_RAMPGENERATOR
END_METHOD

METHOD CALL_OUTPUT
END_METHOD

METHOD CALL_RESETCOMMANDS
END_METHOD

METHOD CALL_RESETOUTPUT
END_METHOD

METHOD CALL_STATEMACHINE
END_METHOD

(* ---- L_TW2P_WINDERJOGGING.pou ---- *)
FUNCTION_BLOCK L_TW2P_WINDERJOGGING
VAR_INPUT
	XENABLE : BOOL;
	XJOGLINEPOS : BOOL;
	XJOGLINENEG : BOOL;
	LRSETDIAMETER : LREAL;
	LRJOGLINEACC : LREAL := 10000;
	LRJOGLINEDEC : LREAL := 10000;
	LRJOGLINEVEL : LREAL := 7200;
	LRJOGLINEJERK : LREAL := 100000;
	XMATERIALFEEDING : BOOL := FALSE;
	XFOLLOWERACTIVE : BOOL;
	LRSTARTREELSPEED : LREAL;
END_VAR
VAR_OUTPUT
	XERROR : BOOL;
	EERRORID : WORD;
	XBUSY : BOOL;
	XDONE : BOOL;
	XENABLESPEEDFOLLOWER : BOOL;
	LRSETREELSPEED : LREAL;
END_VAR
VAR
	XENABLE_OLD : BOOL;
	WSTEPPER : WORD;
	LRVELOCITY : LREAL;
	XMATERIALFEEDING_OLD : BOOL := FALSE;
	L_D94A_SDRAMPGENERATOR1 : L_MC1P_RampGenerator;
END_VAR
END_FUNCTION_BLOCK

METHOD CALL_FB
END_METHOD

METHOD CALL_STATEMACHINE
END_METHOD

METHOD CALL_S001_INIT
END_METHOD

METHOD CALL_S002_READY
END_METHOD

METHOD CALL_S011_JOGPOS
END_METHOD

METHOD CALL_S012_JOGNEG
END_METHOD

METHOD S001_INIT
END_METHOD

METHOD S002_READY
END_METHOD

METHOD S011_JOGPOS
END_METHOD

METHOD S012_JOGNEG
END_METHOD

(* ---- L_TW2P_WINDERSYNCHRONISELINE.pou ---- *)
FUNCTION_BLOCK L_TW2P_WINDERSYNCHRONISELINE
VAR_INPUT
	XENABLE : BOOL;
	XSYNCLINEVEL : BOOL;
	XLOADSTARTREELSPEED : BOOL;
	LRSTARTREELSPEED : LREAL;
	LRGROUNDREELSPEED : LREAL;
	LRCYCLINEVEL : LREAL := 0;
	LRSETDIAMETER : LREAL;
	LRACC : LREAL := 1000;
	LRDEC : LREAL := 1000;
	LRJERK : LREAL := 100000;
	XMATERIALFEEDING : BOOL := FALSE;
END_VAR
VAR_OUTPUT
	XERROR : BOOL;
	EERRORID : WORD;
	XBUSY : BOOL;
	XSYNCHRONISED : BOOL;
	XACCDECSYNC : BOOL;
	LRSETREELSPEEDOUT : LREAL;
END_VAR
VAR
	WSTATE : WORD;
	LRREELSPEEDOUT_INT : LREAL;
	FB_RAMPGENERATOR1 : L_MC1P_RampGenerator;
	XENABLE_OLD : BOOL;
	XMATERIALFEEDING_OLD : BOOL;
	LRSCALEFAKTOR : LREAL;
	LRSCALEFAKTORABS : LREAL;
	WPARMODE : WORD;
	XTMP : BOOL;
END_VAR
END_FUNCTION_BLOCK

METHOD CALL_ERRORHANDLER
END_METHOD

METHOD CALL_FBMETHODS
END_METHOD

METHOD CALL_FB_RAMPGENERATOR
END_METHOD

METHOD CALL_OUTPUT
END_METHOD

METHOD CALL_RESETCOMMANDS
END_METHOD

METHOD CALL_RESETOUTPUT
END_METHOD

METHOD CALL_SETPARMODE
END_METHOD

METHOD CALL_STATEMACHINE
END_METHOD

(* ---- L_TW2P_WINDERTENSIONCTRLSTATE.pou ---- *)
FUNCTION_BLOCK L_TW2P_WINDERTENSIONCTRLSTATE EXTENDS L_TW2P_Winder
VAR_INPUT
	XENABLE : BOOL;
	XENABLEOPERATION : BOOL;
	XRESETERROR : BOOL;
	XQSPAPPLICATION : BOOL;
	XABORT : BOOL;
	XJOGPOS : BOOL;
	XJOGNEG : BOOL;
	XHOMEEXECUTE : BOOL;
	LROVERRIDE : LREAL := 1;
	SCCTRLBASICMOTION : L_TB2P_scCtrlBasicMotion;
	SCPAR : L_TW2P_scPar_WinderTensionCtrlState;
	SCACCESSPOINTS : L_TW2P_scAP_WinderTensionCtrlState;
	XMATERIALFEEDING : BOOL;
	XWINDINGDIRECTION : BOOL;
	XWINDINGDIRECTIONSTANDSTILL : BOOL;
	XJOGLINEPOS : BOOL;
	XJOGLINENEG : BOOL;
	LRSETLINEVEL : LREAL;
	LRSETLINEVELDIAMCALC : LREAL;
	XLOADDIAM : BOOL;
	LRLOADDIAM : LREAL;
	XHOLDDIAM : BOOL;
	XDIAMCALCREDUCED : BOOL;
	XWEBBREAKMONIT : BOOL;
	XSYNCIN : BOOL;
	XTENSCURVE : BOOL;
	XTENSCTRL : BOOL;
	LRSETTENS : LREAL;
	LRACTTENSIN : LREAL;
	LRCTRLINFLUENCESCALED : LREAL;
	XRESETPICTRL : BOOL;
	XRESETICTRL : BOOL;
	XFRICCMPS : BOOL;
	LRSETFRICADAPT : LREAL := 1;
	XEXECUTEIDENTFRIC : BOOL;
	XACCCMPS : BOOL;
	LRMINERTIAADAPT : LREAL := 1;
	XEXECUTEIDENTMINERTIA : BOOL;
	XADAPTSPDCTRLGAIN : BOOL;
	LRADAPTSPDCTRLGAINFACTOR : LREAL := 1;
	XSETMATERIALCOUNTER : BOOL;
	MATERIALCOUNTERVALUES : L_MC1P_IAXIS_REF_MASTERVALUES;
END_VAR
VAR_OUTPUT
	XREADYFOROPERATION : BOOL;
	XOPERATIONENABLED : BOOL;
	XREADYFORMOTION : BOOL;
	XERROR : BOOL;
	XWARNING : BOOL;
	EERRORID : L_IE1P_Error;
	XSTOACTIVE : BOOL;
	XQSPACTIVE : BOOL;
	XABORTBUSY : BOOL;
	XABORTDONE : BOOL;
	XJOGGINGBUSY : BOOL;
	XHOMINGBUSY : BOOL;
	XHOMINGDONE : BOOL;
	XISHOMED : BOOL;
	ETMSTATE : L_TB2P_States := L_TB2P_States.DISABLED;
	SCSTATUSBASICMOTION : L_TB2P_scStatusBasicMotion;
	LRACTVEL : LREAL;
	LRSETVELOUT : LREAL;
	LRACTPOS : LREAL;
	LRSETPOSOUT : LREAL;
	LRACTFOLLOWINGERROR : LREAL;
	SCSIGNALFLOW : L_TW2P_scSF_WinderTensionCtrlState;
	XHOLDDIAMACTIVE : BOOL;
	XDIAMMAX : BOOL;
	XDIAMMIN : BOOL;
	LRSETDIAMOUT : LREAL;
	XWEBBREAK : BOOL;
	XSYNCHRONISED : BOOL;
	XACCDECSYNC : BOOL;
	XWINDINGBUSY : BOOL;
	XUNWIND : BOOL;
	XCONSTANTTENSION : BOOL;
	XTENSINTARGET : BOOL;
	XWNDSPDLIMIT : BOOL;
	LRSETMINERTIAOUT : LREAL;
	XIDENTBUSY : BOOL;
	XIDENTDONE : BOOL;
	LRIDENTMINERTIA : LREAL;
	LRSETSPDCTRLGAINADAPTOUT : LREAL;
	LRMATERIALCOUNTER : LREAL;
	LRLIMITLINEVEL : LREAL;
	XVELOCITYMASTERBUSY : BOOL;
	LRSETLINEVELOUT : LREAL;
	XLINESTOP : BOOL;
END_VAR
VAR_IN_OUT
	AXIS : AXIS_REF;
	PERSISTENTVAR : L_TW2P_PersistentVarWinder;
	ALRFRICTIONCURVE1 : ARRAY [1..66] OF LREAL;
	ALRFRICTIONCURVE2 : ARRAY [1..66] OF LREAL;
	ALRFRICTIONCURVE3 : ARRAY [1..66] OF LREAL;
	ALRFRICTIONCURVE4 : ARRAY [1..66] OF LREAL;
END_VAR
VAR
	TM_INT : L_TW2P_TM_WinderTensionCtrlState := STRUCT(ModuleHandler := ModuleHandler);
	_UICALLMFUNIDXINPUT : UINT := 1;
	_UICALLMFUNIDXOUTPUT : UINT := 1;
	_ASCINPUT : ARRAY [1.._MCCall.c_BufferDepthInput] OF L_TW2P_WinderTensionCtrlStateIn;
	_ASCOUTPUT : ARRAY [1.._MCCall.c_BufferDepthOutput] OF L_TW2P_WinderTensionCtrlStateOut;
	_ASCPARCORE : ARRAY [1.._MCCall.c_BufferDepthInput] OF L_TW2P_scPar_WinderTensionCtrlState;
	_MCCALL : L_UM1P_MCCall;
	_ASCACCESSPOINTSCORE : ARRAY [1.._MCCall.c_BufferDepthInput] OF L_TW2P_scAP_WinderTensionCtrlState;
	_ASCSIGNALFLOWCORE : ARRAY [1.._MCCall.c_BufferDepthOutput] OF L_TW2P_scSF_WinderTensionCtrlState;
	SCPAR_INT : L_TW2P_scPar_WinderTensionCtrlState;
	_SCINPUTVISU : L_TW2P_WinderTensionCtrlStateIn;
	_PSCINPUTVISU : POINTER TO L_TW2P_WinderTensionCtrlStateIn := ADR(_scInputVisu);
	_PSCOUTPUTVISU : POINTER TO L_TW2P_WinderTensionCtrlStateOut := ADR(_ascOutput[1]);
	_PSCPARVISU : POINTER TO L_TW2P_scPar_WinderTensionCtrlState := ADR(scPar_int);
	ITFITECHMODULEINTERNAL : L_TB2P_ITechModuleInternal;
	LRJERKDEC : LREAL;
	LRJOGGINGJERKDEC : LREAL;
	REMAININGTIMEOFPROFILE : LREAL;
	REMAININGTIMEOFPROFILEAVAILABLE : BOOL;
END_VAR
END_FUNCTION_BLOCK

METHOD CALL_COUPLINGREELSPEEDLIMIT
END_METHOD

METHOD CALL_DECOUPLINGREELSPEEDLIMIT
END_METHOD

METHOD GET_ESTATE : L_TB2P_States
END_METHOD

METHOD GET_ETMSTATE : L_TB2P_States
END_METHOD

METHOD GET_LRACTACCTRQ : LREAL
END_METHOD

METHOD GET_LRACTFRICTRQ : LREAL
END_METHOD

METHOD GET_LRACTMOTORTORQUE : LREAL
END_METHOD

METHOD GET_LRACTTENSTRQ : LREAL
END_METHOD

METHOD GET_LRCALCDIAMDIST : LREAL
END_METHOD

METHOD GET_LRCALCDIAMLINESPEED : LREAL
END_METHOD

METHOD GET_LRCALCDIAMREELSPEED : LREAL
END_METHOD

METHOD GET_LRFEEDCONSTANT : LREAL
END_METHOD

METHOD GET_LRLOWERSPEEDLIMIT : LREAL
END_METHOD

METHOD GET_LRMOTORTORQUEREF : LREAL
END_METHOD

METHOD GET_LRRAMPGENOUT : LREAL
END_METHOD

METHOD GET_LRREELSPEEDREF : LREAL
END_METHOD

METHOD GET_LRSETMOTORTORQUE : LREAL
END_METHOD

METHOD GET_LRSETSPEEDCTRLGAINADAPT : LREAL
END_METHOD

METHOD GET_LRSETTOTALTORQUE : LREAL
END_METHOD

METHOD GET_LRSPEEDLOWERLIMIT : LREAL
END_METHOD

METHOD GET_LRSPEEDUPPERLIMIT : LREAL
END_METHOD

METHOD GET_LRTASKCYCLE : LREAL
END_METHOD

METHOD GET_LRTENSCTRLOUT : LREAL
END_METHOD

METHOD GET_LRTENSCURVEOUT : LREAL
END_METHOD

METHOD GET_LRUPPERSPEEDLIMIT : LREAL
END_METHOD

METHOD GET_LRVARMINERTIASCALED : LREAL
END_METHOD

METHOD GET_LRWINDERTORQUEREF : LREAL
END_METHOD

METHOD GET_XCOMMUNICATION : BOOL
END_METHOD

METHOD GET_XDIAMWEBBREAKENABLE : BOOL
VAR_OUTPUT
	XUNIDIRECT : BOOL;
	XUNWINDACTIVE : BOOL;
END_VAR
END_METHOD

METHOD SET_ALRPROCESSCTRLXVALUES
VAR_INPUT
	ALRPROCESSCTRLXVALUES : ARRAY [1..5] OF LREAL;
END_VAR
END_METHOD

METHOD SET_ALRPROCESSCTRLYVALUES
VAR_INPUT
	ALRPROCESSCTRLYVALUES : ARRAY [1..5] OF LREAL;
END_VAR
END_METHOD

METHOD SET_ESTATE
VAR_INPUT
	IN : L_TB2P_States;
END_VAR
END_METHOD

METHOD SET_LRFEEDCONSTANT
VAR_INPUT
	LRIN : LREAL := 0;
END_VAR
END_METHOD

METHOD SET_LRPICTRLINTVALUE
VAR_INPUT
	LRIN : LREAL := 0;
END_VAR
END_METHOD

METHOD SET_LRPROCESSCTRLACC
VAR_INPUT
	LRPROCESSCTRLACC : LREAL := 0.0;
END_VAR
END_METHOD

METHOD SET_LRPROCESSCTRLDEC
VAR_INPUT
	LRPROCESSCTRLDEC : LREAL := 0.0;
END_VAR
END_METHOD

METHOD SET_LRPROCESSCTRLGAINADAPT
VAR_INPUT
	LRPROCESSCTRLGAINADAPT : LREAL := 1;
END_VAR
END_METHOD

METHOD SET_LRPROCESSCTRLINTVALUE
VAR_INPUT
	LRPROCESSCTRLINTVALUE : LREAL := 0.0;
END_VAR
END_METHOD

METHOD SET_LRPROCESSCTRLREDGAIN
VAR_INPUT
	LRPROCESSCTRLREDGAIN : LREAL := 0.0;
END_VAR
END_METHOD

METHOD SET_LRPROCESSCTRLREDRANGE
VAR_INPUT
	LRPROCESSCTRLREDRANGE : LREAL := 0.0;
END_VAR
END_METHOD

METHOD SET_LRREFERENCEMOTORTORQUE
VAR_INPUT
	LRIN : LREAL := 0;
END_VAR
END_METHOD

METHOD SET_LRREFERENCEREELSPEED
VAR_INPUT
	LRIN : LREAL := 0;
END_VAR
END_METHOD

METHOD SET_LRSPEEDOFFSET
VAR_INPUT
	LRIN : LREAL := 0;
END_VAR
END_METHOD

METHOD SET_LRTORQUEOFFSET
VAR_INPUT
	LRIN : LREAL := 0;
END_VAR
END_METHOD

METHOD SET_RPROCESSCTRLDELAYTIME
VAR_INPUT
	RPROCESSCTRLDELAYTIME : REAL := 0.0;
END_VAR
END_METHOD

METHOD SET_RPROCESSCTRLRATEDTIME
VAR_INPUT
	RPROCESSCTRLRATEDTIME : REAL := 0.0;
END_VAR
END_METHOD

METHOD SET_XPICTRLLOADINTVALUE
VAR_INPUT
	XIN : BOOL := FALSE;
END_VAR
END_METHOD

METHOD SET_XPROCESSCTRLLOADINTVALUE
VAR_INPUT
	XPROCESSCTRLLOADINTVALUE : BOOL := FALSE;
END_VAR
END_METHOD

METHOD SET_XSPEEDLIMITENABLEDEXT
VAR_INPUT
	XIN : BOOL := TRUE;
END_VAR
END_METHOD

METHOD SET_XWEBBREAK
VAR_INPUT
	XIN : BOOL := FALSE;
END_VAR
END_METHOD

METHOD CALLFUNCTION
VAR_INPUT
	UIINPUTDATAIDX : UINT;
	UIOUTPUTDATAIDX : UINT;
END_VAR
END_METHOD

METHOD COPYINPUTS : BOOL
VAR_INPUT
	IDX : WORD;
END_VAR
END_METHOD

METHOD COPYOUTPUTS : BOOL
VAR_INPUT
	IDX : WORD;
END_VAR
END_METHOD

METHOD FUNCTIONWASCALLEDTWICE : BOOL
VAR_INPUT
	IDX : WORD;
END_VAR
END_METHOD

METHOD HANDLESTANDARDCALL : BOOL
END_METHOD

METHOD SYNCOUTPUTS
VAR_INPUT
	UICOPYOUTPUTFROMIDX : UINT;
	UICOPYOUTPUTTOIDX : UINT;
END_VAR
END_METHOD

METHOD CALL_INTERNALCTRL
END_METHOD

METHOD GET_PAP : POINTER TO L_TB2P_scAP_TM_MotionControl
END_METHOD

METHOD GET_PPAR : POINTER TO L_TB2P.L_TB2P_scPar_TM_MotionControl
END_METHOD

METHOD GET_PSF : POINTER TO L_TB2P_scSF_TM_MotionControl
END_METHOD

(* ---- L_TW2P_WINDERVELOCITYMASTER.pou ---- *)
FUNCTION_BLOCK L_TW2P_WINDERVELOCITYMASTER
VAR_INPUT
	XENABLE : BOOL;
	XSYNCVEL : BOOL;
	XWINDINGDIRECTION : BOOL;
	LRTASKCYCLETIME : LREAL := 0.001;
	LRSETLINEVEL : LREAL := 0;
	LRACC : LREAL := 1000;
	LRDEC : LREAL := 1000;
	LRJERK : LREAL := 100000;
	XSYNCOUTATTARGET : BOOL;
	LRCYCMATERIALPOS : LREAL;
	LRTARGETMATERIALPOS : LREAL;
	XSETMATERIALCOUNTER : BOOL;
END_VAR
VAR_OUTPUT
	XERROR : BOOL;
	EERRORID : WORD;
	XBUSY : BOOL;
	XSYNCHRONISED : BOOL;
	XACCDECSYNC : BOOL;
	LRSETLINEVELOUT : LREAL;
	LRSETLINEACCOUT : LREAL;
	LRTARGETMATERIALPOSSTOPLINE : LREAL;
	XLINESTOPACTIVE : BOOL;
	LRDISTTOLINESTOP : LREAL;
	XINVALIDSTOPCONDITIONS : BOOL;
END_VAR
VAR
	FB_RAMPGENERATOR1 : L_MC1P_RampGenerator;
	FB_PROFGENERATOR1 : L_MC1P_ProfileGenerator;
	XVELMODE : BOOL;
	XENABLE_OLD : BOOL;
	XSYNCVEL_OLD : BOOL;
	XSETMATERIALCOUNTER_OLD : BOOL;
	LRSETLINEVEL_WNDDIRECTION : LREAL;
	LRSETLINEACC_WNDDIRECTION : LREAL;
	LRDISTTOLINESTOP_OLD : LREAL;
	LRSTOPDIST : LREAL;
	XLINESTOPACTIVENEXTCYLE : BOOL;
	XSYNCOUTATTARGET_LOCK : BOOL;
	XLINESTOPACTIVE_LOCK : BOOL;
	LRTARGETMATERIALPOS_LOCK : LREAL;
	LRDISTTOTARGET_INT : LREAL;
	LRCYCMATERIALPOS_OLD : LREAL;
	LRPGSETVELOUT : LREAL;
	XUSECALCPGSETVELOUT : BOOL := TRUE;
END_VAR
END_FUNCTION_BLOCK

METHOD CALL_ERRORHANDLER
END_METHOD

METHOD CALL_FBMETHODS
END_METHOD

METHOD CALL_OUTPUT
END_METHOD

METHOD CALL_RESETCOMMANDS
END_METHOD

METHOD CALL_RESETOUTPUT
END_METHOD

METHOD CALL_STOPATTARGET
END_METHOD

METHOD GET_LANDERECHNER : LREAL
VAR_INPUT
	LRMATERIALCOUNTER : LREAL;
	LRSETVEL : LREAL;
	LRSETACC : LREAL;
	LRSTOPDEC : LREAL;
	LRSTOPJERK : LREAL;
END_VAR
VAR_OUTPUT
	LRSTOPDIST : LREAL;
	LRSTOPTIME : LREAL;
END_VAR
END_METHOD

METHOD SETLINESTOPACTIVE : BOOL
END_METHOD
